                           IF (#temp16ParameterCMAddress <> 255) AND (#temp16ParameterCMAddress >= #NUMBER_OF_CONTROLMODULES_MIN) AND (#temp16ParameterCMAddress <= #NUMBER_OF_CONTROLMODULES)
                               AND (#temp16ParameterType >= #TYPE_NONE) AND (#temp16ParameterType <= #TYPE_STRING) THEN
                               #temp16TempInt1 := #temp16ParameterCMAddress / 32;    //DWORD - Adress
                               #temp16TempInt2 := #temp16ParameterCMAddress MOD 32;  //Bit - Adress
                               //If parameter is forced (FRC) --> Parameter is used
                               IF (((#tempUsed[#temp16TempInt1] AND SHL(IN := #temp32TempDword1, N := INT_TO_UINT(#temp16TempInt2))) <> 0) = TRUE) THEN
                                   CASE #temp16ParameterType OF
                                           // Check of mode is done in satellite blocks
                                       #TYPE_ANALOG:
                                           REGION Analog
                                               //Bit Masking funtionality for calculate the used Analog parameter and Position of the Parameter name in the HMI Text List 
                                               #ProcessInValueType.IndexAnalog := #ProcessInValueType.IndexAnalog OR SHL(IN := #temp32TempDword1, N := INT_TO_UINT(#temp16IndexOfDefinitionProcessIn));
                                               #ProcessInValueType.NameIndexAnalog := #ProcessInValueType.NameIndexAnalog OR SHL(IN := #temp32TempDword1, N := INT_TO_UINT(#temp16IndexOfDefinition));
                                               IF ((#temp16IndexIO >= #PROCESS_VALUES_IN_MIN) AND (#temp16IndexIO <= #PROCESS_VALUES_IN_ANALOG_MAX)) THEN
                                                   //WinCC Parameter View Faceplate logic
                                                   #ProcessInAna[#temp16IndexAnalog].WQC := #ProcessValueInAnalog[#temp16IndexMTP].WQC;
                                                   #ProcessInAna[#temp16IndexAnalog].OSLevel := #ProcessValueInAnalog[#temp16IndexMTP].OSLevel;
                                                   #ProcessInAna[#temp16IndexAnalog].V := #ProcessValueInAnalog[#temp16IndexMTP].V;
                                                   #ProcessInAna[#temp16IndexAnalog].VQC := #ProcessValueInAnalog[#temp16IndexMTP].VQC;
                                                   #ProcessInAna[#temp16IndexAnalog].SclMinCur := #ProcessValueInAnalog[#temp16IndexMTP].SclMinCur;
                                                   #ProcessInAna[#temp16IndexAnalog].SclMaxCur := #ProcessValueInAnalog[#temp16IndexMTP].SclMaxCur;
                                                   #ProcessInAna[#temp16IndexAnalog].UnitCur := #ProcessValueInAnalog[#temp16IndexMTP].UnitCur;
                                                   #ProcessInAna[#temp16IndexAnalog].SclMinExt := #ProcessValueInAnalog[#temp16IndexMTP].SclMinExt;
                                                   #ProcessInAna[#temp16IndexAnalog].SclMaxExt := #ProcessValueInAnalog[#temp16IndexMTP].SclMaxExt;
                                                   #ProcessInAna[#temp16IndexAnalog].UnitExt := #ProcessValueInAnalog[#temp16IndexMTP].UnitExt;
                                                   #ProcessInAna[#temp16IndexAnalog].Apply := #ProcessValueInAnalog[#temp16IndexMTP].Apply;
                                                   #ProcessInAna[#temp16IndexAnalog].ApplyEn := #ProcessValueInAnalog[#temp16IndexMTP].ApplyEn;
                                               END_IF;
                                               #temp16IndexAnalog := #temp16IndexAnalog + 1;
                                           END_REGION
                                       #TYPE_DIGITAL:
                                           REGION Digital
                                               //Bit Masking funtionality for calculate the used Digital parameter and Position of the Parameter name in the HMI Text List 
                                               #ProcessInValueType.IndexDigital := #ProcessInValueType.IndexDigital OR SHL(IN := #temp32TempDword1, N := INT_TO_UINT(#temp16IndexOfDefinitionProcessIn));
                                               #ProcessInValueType.NameIndexDigital := #ProcessInValueType.NameIndexDigital OR SHL(IN := #temp32TempDword1, N := INT_TO_UINT(#temp16IndexOfDefinition));
                                               IF ((#temp16IndexIO >= #PROCESS_VALUES_IN_MIN) AND (#temp16IndexIO <= #PROCESS_VALUES_IN_DIGITAL_MAX)) THEN
                                                   //WinCC Parameter View Faceplate logic
                                                   #ProcessInDint[#temp16IndexDigital].WQC := #ProcessValueInDigital[#temp16IndexMTP].WQC;
                                                   #ProcessInDint[#temp16IndexDigital].OSLevel := #ProcessValueInDigital[#temp16IndexMTP].OSLevel;
                                                   #ProcessInDint[#temp16IndexDigital].V := #ProcessValueInDigital[#temp16IndexMTP].V;
                                                   #ProcessInDint[#temp16IndexDigital].VQC := #ProcessValueInDigital[#temp16IndexMTP].VQC;
                                                   #ProcessInDint[#temp16IndexDigital].SclMinCur := #ProcessValueInDigital[#temp16IndexMTP].SclMinCur;
                                                   #ProcessInDint[#temp16IndexDigital].SclMaxCur := #ProcessValueInDigital[#temp16IndexMTP].SclMaxCur;
                                                   #ProcessInDint[#temp16IndexDigital].UnitCur := #ProcessValueInDigital[#temp16IndexMTP].UnitCur;
                                                   #ProcessInDint[#temp16IndexDigital].SclMinExt := #ProcessValueInDigital[#temp16IndexMTP].SclMinExt;
                                                   #ProcessInDint[#temp16IndexDigital].SclMaxExt := #ProcessValueInDigital[#temp16IndexMTP].SclMaxExt;
                                                   #ProcessInDint[#temp16IndexDigital].UnitExt := #ProcessValueInDigital[#temp16IndexMTP].UnitExt;
                                                   #ProcessInDint[#temp16IndexDigital].Apply := #ProcessValueInDigital[#temp16IndexMTP].Apply;
                                                   #ProcessInDint[#temp16IndexDigital].ApplyEn := #ProcessValueInDigital[#temp16IndexMTP].ApplyEn;
                                               END_IF;
                                               #temp16IndexDigital := #temp16IndexDigital + 1;
                                           END_REGION
                                       #TYPE_BINARY:
                                           REGION Binary
                                               //Bit Masking funtionality for calculate the used Binary parameter and Position of the Parameter name in the HMI Text List 
                                               #ProcessInValueType.IndexBinary := #ProcessInValueType.IndexBinary OR SHL(IN := #temp32TempDword1, N := INT_TO_UINT(#temp16IndexOfDefinitionProcessIn));
                                               #ProcessInValueType.NameIndexBinary := #ProcessInValueType.NameIndexBinary OR SHL(IN := #temp32TempDword1, N := INT_TO_UINT(#temp16IndexOfDefinition));
                                               IF ((#temp16IndexIO >= #PROCESS_VALUES_IN_MIN) AND (#temp16IndexIO <= #PROCESS_VALUES_IN_BINARY_MAX)) THEN
                                                   //WinCC Parameter View Faceplate logic
                                                   #ProcessInBin[#temp16IndexBinary].WQC := #ProcessValueInBinary[#temp16IndexMTP].WQC;
                                                   #ProcessInBin[#temp16IndexBinary].V := #ProcessValueInBinary[#temp16IndexMTP].V;
                                                   #ProcessInBin[#temp16IndexBinary].VQC := #ProcessValueInBinary[#temp16IndexMTP].VQC;
                                                   #ProcessInBin[#temp16IndexBinary].VState0 := #ProcessValueInBinary[#temp16IndexMTP].VState0;
                                                   #ProcessInBin[#temp16IndexBinary].VState1 := #ProcessValueInBinary[#temp16IndexMTP].VState1;
                                               END_IF;
                                               #temp16IndexBinary := #temp16IndexBinary + 1;
                                           END_REGION
                                       #TYPE_STRING:
                                           REGION String
                                               //Bit Masking funtionality for calculate the used String parameter and Position of the Parameter name in the HMI Text List 
                                               #ProcessInValueType.IndexString := #ProcessInValueType.IndexString OR SHL(IN := #temp32TempDword1, N := INT_TO_UINT(#temp16IndexOfDefinitionProcessIn));
                                               #ProcessInValueType.NameIndexString := #ProcessInValueType.NameIndexString OR SHL(IN := #temp32TempDword1, N := INT_TO_UINT(#temp16IndexOfDefinition));
                                               IF ((#temp16IndexIO >= #PROCESS_VALUES_IN_MIN) AND (#temp16IndexIO <= #PROCESS_VALUES_IN_STRING_MAX)) THEN
                                                   //WinCC Parameter View Faceplate logic
                                                   #ProcessInString[#temp16IndexString].WQC := #ProcessValueInString[#temp16IndexMTP].WQC;
                                                   #ProcessInString[#temp16IndexString].V := #ProcessValueInString[#temp16IndexMTP].V;
                                                   #ProcessInString[#temp16IndexString].VQC := #ProcessValueInString[#temp16IndexMTP].VQC;
                                               END_IF;
                                               #temp16IndexString := #temp16IndexString + 1;
                                           END_REGION
                                   END_CASE;
                               END_IF;
                           END_IF;
                           #temp16IndexOfDefinitionProcessIn := #temp16IndexOfDefinitionProcessIn + 1;
                       END_IF;
                   END_FOR;
               END_IF;
           END_IF;
       END_REGION

       REGION Process Out Values

           REGION Get Start and End index details of the Current /Prepared procedure
               //Current/Prepared procedure selection for parameter display in the faceplate
               //#stat32PrecedureProcessOutMap := -1;
               IF NOT (#ProcessOutValueType.ProcedureReqCurInd) THEN
                   #stat32PrecedureProcessOutMap := #tempSetup.procedure.procedure[#stat16ProceCurIndex].ProcedureProcessOutMap[0];
               ELSIF (#ProcessOutValueType.ProcedureReqCurInd) THEN
                   #stat32PrecedureProcessOutMap := #tempSetup.procedure.procedure[#stat16ProceReqIndex].ProcedureProcessOutMap[0];
               END_IF;
           END_REGION
           //Initialize the used variable values          
           #temp32TempDword1 := 16#1;
           #temp16IndexAnalog := 16#0;
           #temp16IndexDigital := 16#0;
           #temp16IndexBinary := 16#0;
           #temp16IndexString := 16#0;
           //Initialize the Process Out Value index and Name index while changing of Procedure and changing of screen selection b/w Prepared and Current procedure
           IF ((#statLasProcedureCur <> #ProcedureCur) OR (#statLasProcedureReq <> #ProcedureReq) OR (#StatLastProceselProcessOut <> #ProcessOutValueType.ProcedureReqCurInd)
               OR (((#ProcedureCur = 16#0) AND NOT #ProcessOutValueType.ProcedureReqCurInd) OR ((#ProcedureReq = 16#0) AND #ProcessOutValueType.ProcedureReqCurInd))) THEN
               #ProcessOutValueType.IndexAnalog := 16#0;
               #ProcessOutValueType.NameIndexAnalog := 16#0;
               #ProcessOutValueType.IndexDigital := 16#0;
               #ProcessOutValueType.NameIndexDigital := 16#0;
               #ProcessOutValueType.IndexBinary := 16#0;
               #ProcessOutValueType.NameIndexBinary := 16#0;
               #ProcessOutValueType.IndexString := 16#0;
               #ProcessOutValueType.NameIndexString := 16#0;
           END_IF;
           //Used/Mapped parameter count with individual parameter type will written from the Tool
           #statTotalProcessOutValues := #MAPPED_PROCESS_OUT_ANALOG + #MAPPED_PROCESS_OUT_DIGITAL + #MAPPED_PROCESS_OUT_BINARY + #MAPPED_PROCESS_OUT_STRING - 1;
           IF (((#ProcedureCur <> 16#0) AND NOT #ProcessOutValueType.ProcedureReqCurInd) OR ((#ProcedureReq <> 16#0) AND #ProcessOutValueType.ProcedureReqCurInd)) THEN
               IF ((#statTotalProcessOutValues >= 0) AND (#statTotalProcessOutValues <= #PROCESS_VALUES_OUT_MAX)) THEN
                   #temp16IndexOfDefinitionProcessOut := 16#0;
                   FOR #temp16IndexOfDefinition := #PROCESS_VALUES_OUT_MIN TO #statTotalProcessOutValues BY 1 DO
                       #temp16ParameterCMAddress := BYTE_TO_INT(#tempSetup.processValueOutData.definition[#temp16IndexOfDefinition].controlModule);
                       #temp16ParameterType := #tempSetup.processValueOutData.definition[#temp16IndexOfDefinition].type;
                       #temp16IndexMTP := #tempSetup.processValueOutData.definition[#temp16IndexOfDefinition].indexMTP;
                       #tempUsed := #tempSetup.processValueOutData.used;
                       // Find the procedure information assigned with the processOut values
                       IF (((#stat32PrecedureProcessOutMap AND SHL(IN := #temp32TempDword1, N := INT_TO_UINT(#temp16IndexOfDefinition))) <> 0) = TRUE) THEN
                           #temp16IndexIO := #tempSetup.processValueOutData.definition[#temp16IndexOfDefinition].indexIO;

                           IF (#temp16ParameterCMAddress <> 255) AND (#temp16ParameterCMAddress >= #NUMBER_OF_CONTROLMODULES_MIN) AND (#temp16ParameterCMAddress <= #NUMBER_OF_CONTROLMODULES)
                               AND (#temp16ParameterType >= #TYPE_NONE) AND (#temp16ParameterType <= #TYPE_STRING) THEN
                               #temp16TempInt1 := #temp16ParameterCMAddress / 32;    //DWORD - Adress
                               #temp16TempInt2 := #temp16ParameterCMAddress MOD 32;  //Bit - Adress
                               //If parameter is forced (FRC) --> Parameter is used
                               IF (((#tempUsed[#temp16TempInt1] AND SHL(IN := #temp32TempDword1, N := INT_TO_UINT(#temp16TempInt2))) <> 0) = TRUE) THEN
                                   CASE #temp16ParameterType OF
                                       #TYPE_ANALOG:
                                           REGION Analog
                                               //Bit Masking funtionality for calculate the used Analog parameter and Position of the Parameter name in the HMI Text List                                         
                                               #ProcessOutValueType.IndexAnalog := #ProcessOutValueType.IndexAnalog OR SHL(IN := #temp32TempDword1, N := INT_TO_UINT(#temp16IndexOfDefinitionProcessOut));
                                               #ProcessOutValueType.NameIndexAnalog := #ProcessOutValueType.NameIndexAnalog OR SHL(IN := #temp32TempDword1, N := INT_TO_UINT(#temp16IndexOfDefinition));
                                               IF ((#temp16IndexIO >= #PROCESS_VALUES_OUT_MIN) AND (#temp16IndexIO <= #PROCESS_VALUES_OUT_ANALOG_MAX)) THEN
                                                   //WinCC Parameter View Faceplate logic
                                                   #ProcessOutAna[#temp16IndexAnalog].WQC := #ProcessValueOutAnalog[#temp16IndexMTP].WQC;
                                                   #ProcessOutAna[#temp16IndexAnalog].V := #ProcessValueOutAnalog[#temp16IndexMTP].V;
                                                   #ProcessOutAna[#temp16IndexAnalog].VSclMin := #ProcessValueOutAnalog[#temp16IndexMTP].VSclMin;
                                                   #ProcessOutAna[#temp16IndexAnalog].VSclMax := #ProcessValueOutAnalog[#temp16IndexMTP].VSclMax;
                                                   #ProcessOutAna[#temp16IndexAnalog].VUnit := #ProcessValueOutAnalog[#temp16IndexMTP].VUnit;
                                               END_IF;
                                               #temp16IndexAnalog := #temp16IndexAnalog + 1;
                                           END_REGION
                                       #TYPE_DIGITAL:
                                           REGION Digital
                                               //Bit Masking funtionality for calculate the used Digital parameter and Position of the Parameter name in the HMI Text List                                         
                                               #ProcessOutValueType.IndexDigital := #ProcessOutValueType.IndexDigital OR SHL(IN := #temp32TempDword1, N := INT_TO_UINT(#temp16IndexOfDefinitionProcessOut));
                                               #ProcessOutValueType.NameIndexDigital := #ProcessOutValueType.NameIndexDigital OR SHL(IN := #temp32TempDword1, N := INT_TO_UINT(#temp16IndexOfDefinition));
                                               IF ((#temp16IndexIO >= #PROCESS_VALUES_OUT_MIN) AND (#temp16IndexIO <= #PROCESS_VALUES_OUT_DIGITAL_MAX)) THEN
                                                   //WinCC Parameter View Faceplate logic
                                                   #ProcessOutDint[#temp16IndexDigital].WQC := #ProcessValueOutDigital[#temp16IndexMTP].WQC;
                                                   #ProcessOutDint[#temp16IndexDigital].V := #ProcessValueOutDigital[#temp16IndexMTP].V;
                                                   #ProcessOutDint[#temp16IndexDigital].VSclMin := #ProcessValueOutDigital[#temp16IndexMTP].VSclMin;
                                                   #ProcessOutDint[#temp16IndexDigital].VSclMax := #ProcessValueOutDigital[#temp16IndexMTP].VSclMax;
                                                   #ProcessOutDint[#temp16IndexDigital].VUnit := #ProcessValueOutDigital[#temp16IndexMTP].VUnit;
                                               END_IF;
                                               #temp16IndexDigital := #temp16IndexDigital + 1;
                                           END_REGION
                                       #TYPE_BINARY:
                                           REGION Binary
                                               //Bit Masking funtionality for calculate the used Binary parameter and Position of the Parameter name in the HMI Text List 
                                               #ProcessOutValueType.IndexBinary := #ProcessOutValueType.IndexBinary OR SHL(IN := #temp32TempDword1, N := INT_TO_UINT(#temp16IndexOfDefinitionProcessOut));
                                               #ProcessOutValueType.NameIndexBinary := #ProcessOutValueType.NameIndexBinary OR SHL(IN := #temp32TempDword1, N := INT_TO_UINT(#temp16IndexOfDefinition));
                                               IF ((#temp16IndexIO >= #PROCESS_VALUES_OUT_MIN) AND (#temp16IndexIO <= #PROCESS_VALUES_OUT_BINARY_MAX)) THEN
                                                   //WinCC Parameter View Faceplate logic
                                                   #ProcessOutBin[#temp16IndexBinary].WQC := #ProcessValueOutBinary[#temp16IndexMTP].WQC;
                                                   #ProcessOutBin[#temp16IndexBinary].V := #ProcessValueOutBinary[#temp16IndexMTP].V;
                                                   #ProcessOutBin[#temp16IndexBinary].VState0 := #ProcessValueOutBinary[#temp16IndexMTP].VState0;
                                                   #ProcessOutBin[#temp16IndexBinary].VState1 := #ProcessValueOutBinary[#temp16IndexMTP].VState1;
                                               END_IF;
                                               #temp16IndexBinary := #temp16IndexBinary + 1;
                                           END_REGION
                                       #TYPE_STRING:
                                           REGION String
                                               //Bit Masking funtionality for calculate the used String parameter and Position of the Parameter name in the HMI Text List 
                                               #ProcessOutValueType.IndexString := #ProcessOutValueType.IndexString OR SHL(IN := #temp32TempDword1, N := INT_TO_UINT(#temp16IndexOfDefinitionProcessOut));
                                               #ProcessOutValueType.NameIndexString := #ProcessOutValueType.NameIndexString OR SHL(IN := #temp32TempDword1, N := INT_TO_UINT(#temp16IndexOfDefinition));
                                               IF ((#temp16IndexIO >= #PROCESS_VALUES_OUT_MIN) AND (#temp16IndexIO <= #PROCESS_VALUES_OUT_STRING_MAX)) THEN
                                                   //WinCC Parameter View Faceplate logic
                                                   #ProcessOutString[#temp16IndexString].WQC := #ProcessValueOutString[#temp16IndexMTP].WQC;
                                                   #ProcessOutString[#temp16IndexString].Text := #ProcessValueOutString[#temp16IndexMTP].Text;
                                               END_IF;
                                               #temp16IndexString := #temp16IndexString + 1;
                                           END_REGION
                                   END_CASE;
                               END_IF;
                           END_IF;
                           #temp16IndexOfDefinitionProcessOut := #temp16IndexOfDefinitionProcessOut + 1;
                       END_IF;
                   END_FOR;
               END_IF;
           END_IF;
       END_REGION

       REGION Report Values

           REGION Get Start and End index details of the Current /Prepared procedure
               //Current/Prepared procedure selection for parameter display in the faceplate
              // #stat32PrecedureReportMap := -1;
               IF NOT (#ReportValueType.ProcedureReqCurInd) THEN
                   #stat32PrecedureReportMap := #tempSetup.procedure.procedure[#stat16ProceCurIndex].ProcedureReportMap[0];
               ELSIF (#ReportValueType.ProcedureReqCurInd) THEN
                   #stat32PrecedureReportMap := #tempSetup.procedure.procedure[#stat16ProceReqIndex].ProcedureReportMap[0];
               END_IF;
           END_REGION
           //Initialize the used variable values        
           #temp32TempDword1 := 16#1;
           #temp16IndexAnalog := 16#0;
           #temp16IndexDigital := 16#0;
           #temp16IndexBinary := 16#0;
           #temp16IndexString := 16#0;
           //Initialize the Process Out Value index and Name index while changing of Procedure and changing of screen selection b/w Prepared and Current procedure
           IF ((#statLasProcedureCur <> #ProcedureCur) OR (#statLasProcedureReq <> #ProcedureReq) OR (#StatLastProceselReport <> #ReportValueType.ProcedureReqCurInd)
               OR (((#ProcedureCur = 16#0) AND NOT #ReportValueType.ProcedureReqCurInd) OR ((#ProcedureReq = 16#0) AND #ReportValueType.ProcedureReqCurInd))) THEN
               #ReportValueType.IndexAnalog := 16#0;
               #ReportValueType.NameIndexAnalog := 16#0;
               #ReportValueType.IndexDigital := 16#0;
               #ReportValueType.NameIndexDigital := 16#0;
               #ReportValueType.IndexBinary := 16#0;
               #ReportValueType.NameIndexBinary := 16#0;
               #ReportValueType.IndexString := 16#0;
               #ReportValueType.NameIndexString := 16#0;
           END_IF;
           //Used/Mapped parameter count with individual parameter type will written from the Tool
           #statTotalReportValues := #MAPPED_REPORT_ANALOG + #MAPPED_REPORT_DIGITAL + #MAPPED_REPORT_BINARY + #MAPPED_REPORT_STRING - 1;
           IF (((#ProcedureCur <> 16#0) AND NOT #ReportValueType.ProcedureReqCurInd) OR ((#ProcedureReq <> 16#0) AND #ReportValueType.ProcedureReqCurInd)) THEN
               IF ((#statTotalReportValues >= 0) AND (#statTotalReportValues <= #REPORT_VALUES_MAX)) THEN
                   #temp16IndexOfDefinitionReport := 16#0;
                   FOR #temp16IndexOfDefinition := #REPORT_VALUES_MIN TO #statTotalReportValues BY 1 DO
                       #temp16ParameterCMAddress := BYTE_TO_INT(#tempSetup.reportValueData.definition[#temp16IndexOfDefinition].controlModule);
                       #temp16ParameterType := #tempSetup.reportValueData.definition[#temp16IndexOfDefinition].type;
                       #temp16IndexMTP := #tempSetup.reportValueData.definition[#temp16IndexOfDefinition].indexMTP;
                       #tempUsed := #tempSetup.reportValueData.used;
                       // Find the procedure information assigned with the report values
                       IF (((#stat32PrecedureReportMap AND SHL(IN := #temp32TempDword1, N := INT_TO_UINT(#temp16IndexOfDefinition))) <> 0) = TRUE) THEN
                           #temp16IndexIO := #tempSetup.reportValueData.definition[#temp16IndexOfDefinition].indexIO;

                           IF (#temp16ParameterCMAddress <> 255) AND (#temp16ParameterCMAddress >= #NUMBER_OF_CONTROLMODULES_MIN) AND (#temp16ParameterCMAddress <= #NUMBER_OF_CONTROLMODULES)
                               AND (#temp16ParameterType >= #TYPE_NONE) AND (#temp16ParameterType <= #TYPE_STRING) THEN
                               #temp16TempInt1 := #temp16ParameterCMAddress / 32;    //DWORD - Adress
                               #temp16TempInt2 := #temp16ParameterCMAddress MOD 32;  //Bit - Adress
                               //If parameter is forced (FRC) --> Parameter is used
                               IF (((#tempUsed[#temp16TempInt1] AND SHL(IN := #temp32TempDword1, N := INT_TO_UINT(#temp16TempInt2))) <> 0) = TRUE) THEN
                                   CASE #temp16ParameterType OF
                                       #TYPE_ANALOG:
                                           REGION Analog
                                               //Bit Masking funtionality for calculate the used Analog parameter and Position of the Parameter name in the HMI Text List 
                                               #ReportValueType.IndexAnalog := #ReportValueType.IndexAnalog OR SHL(IN := #temp32TempDword1, N := INT_TO_UINT(#temp16IndexOfDefinitionReport));
                                               #ReportValueType.NameIndexAnalog := #ReportValueType.NameIndexAnalog OR SHL(IN := #temp32TempDword1, N := INT_TO_UINT(#temp16IndexOfDefinition));
                                               IF ((#temp16IndexIO >= #REPORT_VALUES_MIN) AND (#temp16IndexIO <= #REPORT_VALUES_ANALOG_MAX)) THEN
                                                   //WinCC Parameter View Faceplate logic
                                                   #ReportAna[#temp16IndexAnalog].WQC := #ReportValueAnalog[#temp16IndexMTP].WQC;
                                                   #ReportAna[#temp16IndexAnalog].V := #ReportValueAnalog[#temp16IndexMTP].V;
                                                   #ReportAna[#temp16IndexAnalog].VSclMin := #ReportValueAnalog[#temp16IndexMTP].VSclMin;
                                                   #ReportAna[#temp16IndexAnalog].VSclMax := #ReportValueAnalog[#temp16IndexMTP].VSclMax;
                                                   #ReportAna[#temp16IndexAnalog].VUnit := #ReportValueAnalog[#temp16IndexMTP].VUnit;
                                                   #ReportAna[#temp16IndexAnalog].MissedValue := #ReportValueAnalog[#temp16IndexMTP].MissedValue;
                                               END_IF;
                                               #temp16IndexAnalog := #temp16IndexAnalog + 1;
                                           END_REGION
                                       #TYPE_DIGITAL:
                                           REGION Digital
                                               //Bit Masking funtionality for calculate the used Digital parameter and Position of the Parameter name in the HMI Text List 
                                               #ReportValueType.IndexDigital := #ReportValueType.IndexDigital OR SHL(IN := #temp32TempDword1, N := INT_TO_UINT(#temp16IndexOfDefinitionReport));
                                               #ReportValueType.NameIndexDigital := #ReportValueType.NameIndexDigital OR SHL(IN := #temp32TempDword1, N := INT_TO_UINT(#temp16IndexOfDefinition));
                                               IF ((#temp16IndexIO >= #REPORT_VALUES_MIN) AND (#temp16IndexIO <= #REPORT_VALUES_DIGITAL_MAX)) THEN
                                                   //WinCC Parameter View Faceplate logic
                                                   #ReportDint[#temp16IndexDigital].WQC := #ReportValueDigital[#temp16IndexMTP].WQC;
                                                   #ReportDint[#temp16IndexDigital].V := #ReportValueDigital[#temp16IndexMTP].V;
                                                   #ReportDint[#temp16IndexDigital].VSclMin := #ReportValueDigital[#temp16IndexMTP].VSclMin;
                                                   #ReportDint[#temp16IndexDigital].VSclMax := #ReportValueDigital[#temp16IndexMTP].VSclMax;
                                                   #ReportDint[#temp16IndexDigital].VUnit := #ReportValueDigital[#temp16IndexMTP].VUnit;
                                                   #ReportDint[#temp16IndexDigital].MissedValue := #ReportValueDigital[#temp16IndexMTP].MissedValue;
                                               END_IF;
                                               #temp16IndexDigital := #temp16IndexDigital + 1;
                                           END_REGION
                                       #TYPE_BINARY:
                                           REGION Binary
                                               //Bit Masking funtionality for calculate the used Binary parameter and Position of the Parameter name in the HMI Text List 
                                               #ReportValueType.IndexBinary := #ReportValueType.IndexBinary OR SHL(IN := #temp32TempDword1, N := INT_TO_UINT(#temp16IndexOfDefinitionReport));
                                               #ReportValueType.NameIndexBinary := #ReportValueType.NameIndexBinary OR SHL(IN := #temp32TempDword1, N := INT_TO_UINT(#temp16IndexOfDefinition));
                                               IF ((#temp16IndexIO >= #REPORT_VALUES_MIN) AND (#temp16IndexIO <= #REPORT_VALUES_BINARY_MAX)) THEN
                                                   //WinCC Parameter View Faceplate logic
                                                   #ReportBin[#temp16IndexBinary].WQC := #ReportValueBinary[#temp16IndexMTP].WQC;
                                                   #ReportBin[#temp16IndexBinary].V := #ReportValueBinary[#temp16IndexMTP].V;
                                                   #ReportBin[#temp16IndexBinary].VState0 := #ReportValueBinary[#temp16IndexMTP].VState0;
                                                   #ReportBin[#temp16IndexBinary].VState1 := #ReportValueBinary[#temp16IndexMTP].VState1;
                                                   #ReportBin[#temp16IndexBinary].MissedValue := #ReportValueBinary[#temp16IndexMTP].MissedValue;
                                               END_IF;
                                               #temp16IndexBinary := #temp16IndexBinary + 1;
                                           END_REGION
                                       #TYPE_STRING:
                                           REGION String
                                               //Bit Masking funtionality for calculate the used String parameter and Position of the Parameter name in the HMI Text List 
                                               #ReportValueType.IndexString := #ReportValueType.IndexString OR SHL(IN := #temp32TempDword1, N := INT_TO_UINT(#temp16IndexOfDefinitionReport));
                                               #ReportValueType.NameIndexString := #ReportValueType.NameIndexString OR SHL(IN := #temp32TempDword1, N := INT_TO_UINT(#temp16IndexOfDefinition));
                                               IF ((#temp16IndexIO >= #REPORT_VALUES_MIN) AND (#temp16IndexIO <= #REPORT_VALUES_STRING_MAX)) THEN

                                                   //WinCC Parameter View Faceplate logic
                                                   #ReportString[#temp16IndexString].WQC := #ReportValueString[#temp16IndexMTP].WQC;
                                                   #ReportString[#temp16IndexString].Text := #ReportValueString[#temp16IndexMTP].Text;
                                                   #ReportString[#temp16IndexString].MissedValue := #ReportValueString[#temp16IndexMTP].MissedValue;
                                               END_IF;
                                               #temp16IndexString := #temp16IndexString + 1;
                                           END_REGION
                                   END_CASE;
                               END_IF;
                           END_IF;
                           #temp16IndexOfDefinitionReport := #temp16IndexOfDefinitionReport + 1;
                       END_IF;
                   END_FOR;
               END_IF;
           END_IF;
       END_REGION  

       //Move last valid value 
       #statLasProcedureCur := #ProcedureCur;
       #statLasProcedureReq := #ProcedureReq;
       #statLastReqProcedSelected := #ProcedureParaType.ProcedureReqCurInd;
       #StatLastProceselProcessIn := #ProcessInValueType.ProcedureReqCurInd;
       #StatLastProceselProcessOut := #ProcessOutValueType.ProcedureReqCurInd;
       #StatLastProceselReport := #ReportValueType.ProcedureReqCurInd;
END_FUNCTION_BLOCK

FUNCTION_BLOCK "CM_Interface"   // FB5, SCL
{ S7_Optimized_Access := 'TRUE' }
// stored: MemoryReserve 100, SetENOAutomatically false
   VAR_INPUT
      CmCommand { ExternalAccessible := 'False'; ExternalVisible := 'False'; ExternalWritable := 'False'} : Array[0..29] of Bool;
      Procedure_Param { ExternalAccessible := 'False'; ExternalVisible := 'False'; ExternalWritable := 'False'} : Array[0..31] of Real;
      Config_Param : Array[0..31] of Bool;
      ProcessValueIn_Bool : Array[0..31] of Bool;
      ProcessValueIn_Real : Array[0..31] of Real;
      CmFbOnOff { ExternalAccessible := 'False'; ExternalVisible := 'False'; ExternalWritable := 'False'} : Array[0..29] of Bool;
      DosingSpeed : Real;
      Auto_Man : Bool;
      Oos : Bool;
   END_VAR
   VAR_OUTPUT
      CM_P100 { ExternalAccessible := 'False'; ExternalVisible := 'False'; ExternalWritable := 'False'} : "DigVal";
      CM_P101 { ExternalAccessible := 'False'; ExternalVisible := 'False'; ExternalWritable := 'False'} : "DigVal";
      CM_FIC100 { ExternalAccessible := 'False'; ExternalVisible := 'False'; ExternalWritable := 'False'} : "DigVal";
      CM_V100 { ExternalAccessible := 'False'; ExternalVisible := 'False'; ExternalWritable := 'False'} : "DigVal";
      FlowRate { ExternalAccessible := 'False'; ExternalVisible := 'False'; ExternalWritable := 'False'} : "AnaVal";
      Liter { ExternalAccessible := 'False'; ExternalVisible := 'False'; ExternalWritable := 'False'} : "AnaVal";
      ExternalLevel : "AnaVal";
      PEA_inlet_Vlv_opened : "DigVal";
      PVConnected : "DigVal";
   END_VAR
   VAR
      Pos_edge : Bool;
      Neg_edge : Bool;
   END_VAR
   VAR_TEMP
      State : "Service_States";
   END_VAR
BEGIN
   REGION Bool TO DigVal
       //CM Pump 100
       "BoolToDigVal"(In := #CmCommand[0],
                      ST := 16#80,
                      Out => #CM_P100);
       //CM Pump 101
       "BoolToDigVal"(In := #CmCommand[1],
                      ST := 16#80,
                      Out => #CM_P101);
       //CM Controler 100
       "BoolToDigVal"(In := #CmCommand[2],
                      ST := 16#80,
                      Out => #CM_FIC100);
       //CM Valve 100
       "BoolToDigVal"(In := #CmCommand[3],
                      ST := 16#80,
                      Out => #CM_V100);
   END_REGION

   REGION Real TO AnaVal
       //Flow
       "RealToAnaVal"(In := #Procedure_Param[0],
                      ST := 16#80,
                      Out => #FlowRate);
       //Liter
       "RealToAnaVal"(In := #Procedure_Param[1],
                      ST := 16#80,
                      Out => #Liter);
                   END_REGION

   REGION other values
       //Dosing Speed
       "Dose".ProcessValueOutAnalogIn[0] := #DosingSpeed;

       //Configuration parameter
       "BoolToDigVal"(In := #Config_Param[0],
                      ST := 16#80,
                      Out => #PVConnected);
       //process value input
       "RealToAnaVal"(In := #ProcessValueIn_Real[0],
                      ST := 16#80,
                      Out => #ExternalLevel);
       "BoolToDigVal"(In := #ProcessValueIn_Bool[0],
                      ST := 16#80,
                      Out => #PEA_inlet_Vlv_opened);
   END_REGION


   REGION Set auto/man mode & Int/Ext
       //check for positive edge at Dose.Oos
       "R_TRIG_DB"(CLK := #Oos,
                   Q => #Neg_edge);

       //Set POs to auto mode
       IF #Auto_Man = TRUE THEN
           "FIC100_Type".Cmd_Man := FALSE;
           "P100_Type".Cmd_Man := FALSE;
           "V100_Type".Cmd_Man := FALSE;
           "P101_Type".Cmd_Man := FALSE;
           "FIC100_Type".Cmd_Auto := TRUE;
           "P100_Type".Cmd_Auto := TRUE;
           "V100_Type".Cmd_Auto := TRUE;
           "P101_Type".Cmd_Auto := TRUE;
       //Set POs to man mode
       ELSIF #Neg_edge = TRUE THEN
           "FIC100_Type".Cmd_Auto := FALSE;
           "P100_Type".Cmd_Auto := FALSE;
           "V100_Type".Cmd_Auto := FALSE;
           "P101_Type".Cmd_Auto := FALSE;
           "FIC100_Type".Cmd_Man := TRUE;
           "P100_Type".Cmd_Man := TRUE;
           "V100_Type".Cmd_Man := TRUE;
           "P101_Type".Cmd_Man := TRUE;
       //Reset Value
       ELSE
           "FIC100_Type".Cmd_Auto := FALSE;
           "P100_Type".Cmd_Auto := FALSE;
           "V100_Type".Cmd_Auto := FALSE;
           "P101_Type".Cmd_Auto := FALSE;
           "FIC100_Type".Cmd_Man := FALSE;
           "P100_Type".Cmd_Man := FALSE;
           "V100_Type".Cmd_Man := FALSE;
           "P101_Type".Cmd_Man := FALSE;
       END_IF;
   END_REGION
END_FUNCTION_BLOCK

FUNCTION_BLOCK "Service_Command_Logic"   // FB3, SCL
{ S7_Optimized_Access := 'TRUE' }
// stored: MemoryReserve 100, SetENOAutomatically false
   VAR_INPUT
      Level : Real;
      ProcedureID_cur : DWord;
   END_VAR
   VAR_TEMP
      i : Int;
      State : "Service_States";
   END_VAR
BEGIN
   //Set service to hold, if the level of the tank falls under 0,45 during the 
   //procedures DoseByVolume and DoseByFlow
   IF #Level < 45 AND "Dose".Information.state = #State.Execute AND "Dose".MTP.ServiceControl.ProcedureCur <> 3 THEN
       "Dose".CommandForce.hold := TRUE;
       FOR #i := 0 TO 1 BY 1 DO
           "Dose".Procedure[#i].ProcedureEnable.Unhold.ST := 16#80;
           "Dose".Procedure[#i].ProcedureEnable.Unhold.Value := false;
       END_FOR;
   END_IF;
   IF "Dose".Information.state = #State.Held THEN
       "Dose".CommandForce.hold := FALSE;
   END_IF;
   IF "Dose".Information.state = #State.Held AND #Level >= 1.0 THEN
       FOR #i := 0 TO 1 BY 1 DO
           "Dose".Procedure[#i].ProcedureEnable.Unhold.ST := 16#80;
           "Dose".Procedure[#i].ProcedureEnable.Unhold.Value := true;
       END_FOR;
   END_IF;


   //Set service to abort, if the pump is in failure
   IF "P100_Type".GrpErr = True OR "P101_Type".GrpErr THEN
       "Dose".CommandForce.abort := TRUE;
       FOR #i := 0 TO 2 BY 1 DO
           "Dose".Procedure[#i].ProcedureEnable.Start.ST := 16#80;
           "Dose".Procedure[#i].ProcedureEnable.Start.Value := false;
       END_FOR;
   ELSIF ("Dose".Information.state = #State.Aborted OR "Dose".Information.state = #State.Idle) AND ("P100_Type".GrpErr = False OR "P101_Type".GrpErr) THEN
       "Dose".CommandForce.abort := false;
       FOR #i := 0 TO 2 BY 1 DO
           "Dose".Procedure[#i].ProcedureEnable.Start.ST := 16#80;
           "Dose".Procedure[#i].ProcedureEnable.Start.Value := true;
       END_FOR;
   END_IF;
END_FUNCTION_BLOCK

FUNCTION "BoolToDigVal" : Void   // FC10, SCL
{ S7_Optimized_Access := 'TRUE' }
// stored: SetENOAutomatically false
   VAR_INPUT
      In : Bool;
      ST : Byte;
   END_VAR
   VAR_OUTPUT
      Out : "DigVal";
   END_VAR
BEGIN
   #Out.ST := #ST;
   #Out.Value := #In;
END_FUNCTION

FUNCTION "PositionText" : Void   // FC18, SCL
{ S7_Optimized_Access := 'TRUE' }
// stored: SetENOAutomatically false
   VAR_INPUT
      PosID_1 : Bool;
      PosID_2 : Bool;
      PosID_3 : Bool;
      PosID_4 : Bool;
      PosID_5 : Bool;
      PosID_6 : Bool;
      PosID_7 : Bool;
      PosID_8 : Bool;
      PosID_9 : Bool;
      PosID_10 : Bool;
      PosID_0 : Bool;
   END_VAR
BEGIN
   IF #PosID_1 = True THEN
       "Dose".PosTextIDLi := 1;
   ELSIF #PosID_2 = True THEN
       "Dose".PosTextIDLi := 2;
   ELSIF #PosID_3 = True THEN
       "Dose".PosTextIDLi := 3;
   ELSIF #PosID_4 = True THEN
       "Dose".PosTextIDLi := 4;
   ELSIF #PosID_5 = True THEN
       "Dose".PosTextIDLi := 5;
   ELSIF #PosID_6 = True THEN
       "Dose".PosTextIDLi := 6;
   ELSIF #PosID_7 = True THEN
       "Dose".PosTextIDLi := 7;
   ELSIF #PosID_8 = True THEN
       "Dose".PosTextIDLi := 8;
   ELSIF #PosID_9 = True THEN
       "Dose".PosTextIDLi := 9;
   ELSIF #PosID_10 = True THEN
       "Dose".PosTextIDLi := 10;
   ELSIF #PosID_0 = True THEN
       "Dose".PosTextIDLi := 0;
   END_IF;
END_FUNCTION

FUNCTION "FIC100" : Void   // FC5, FBD
{ S7_Optimized_Access := 'TRUE' }
// stored: SetENOAutomatically false
   VAR_TEMP
      Temp : "DigVal";
      State : "Service_States";
      Interlock : "DigVal";
   END_VAR
BEGIN

REGION Network 1: PIDConL interconnections
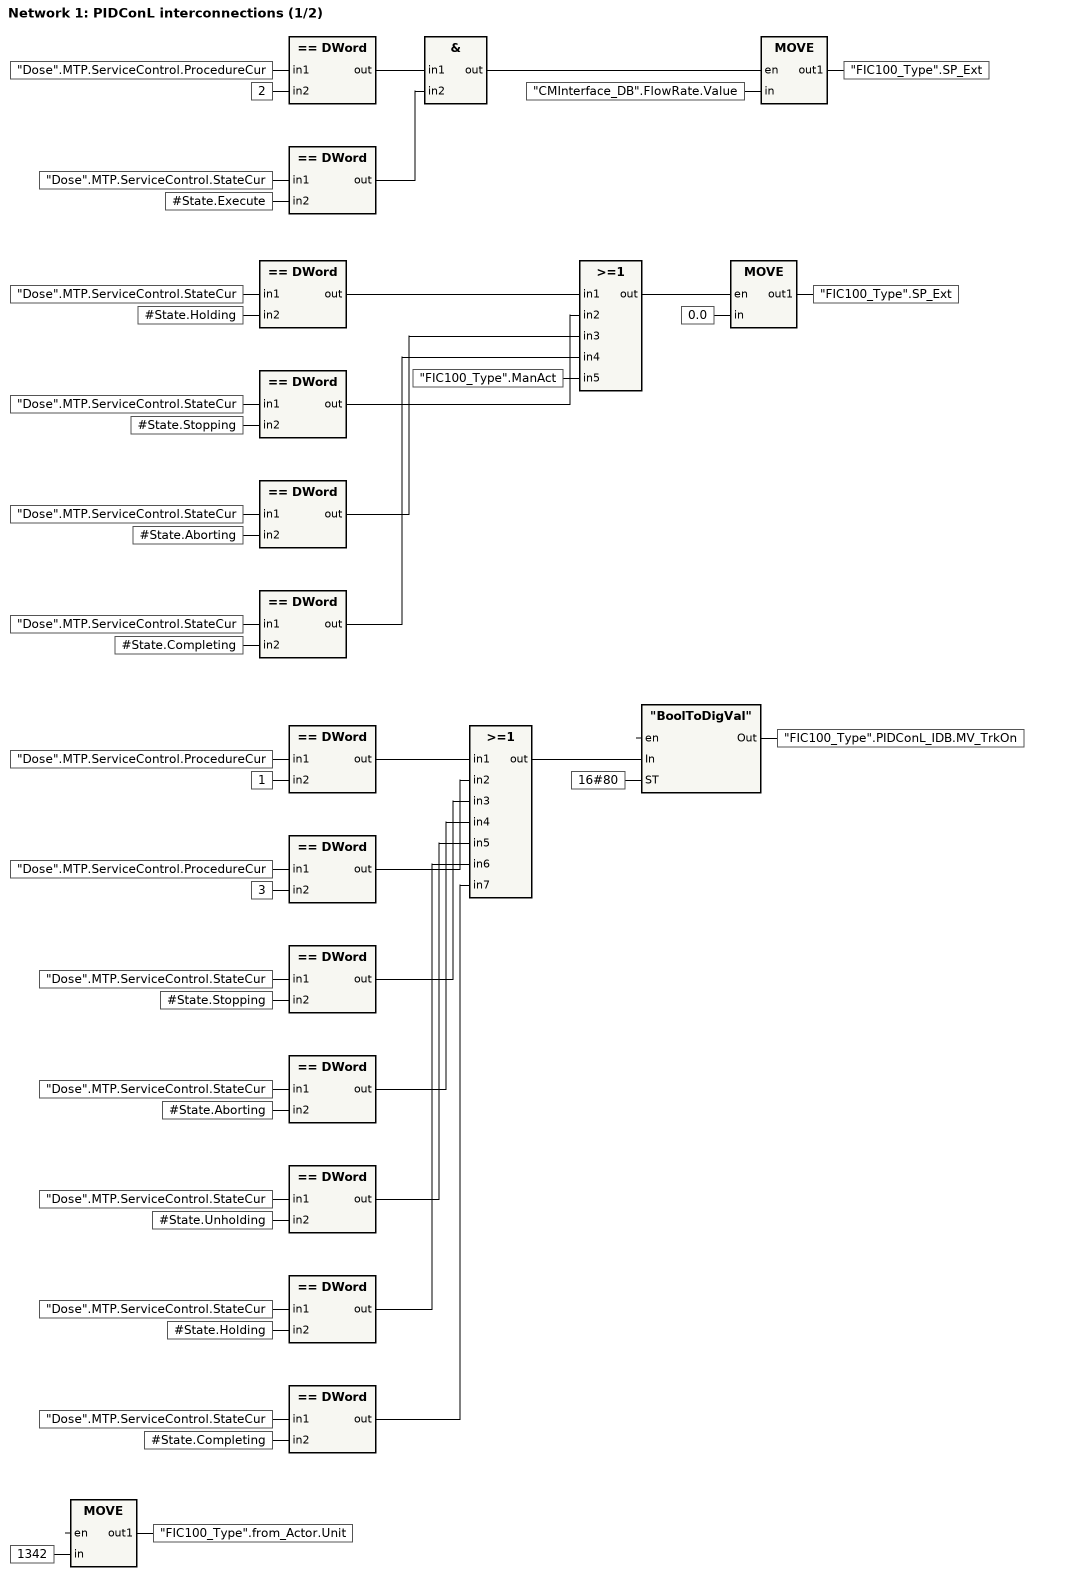
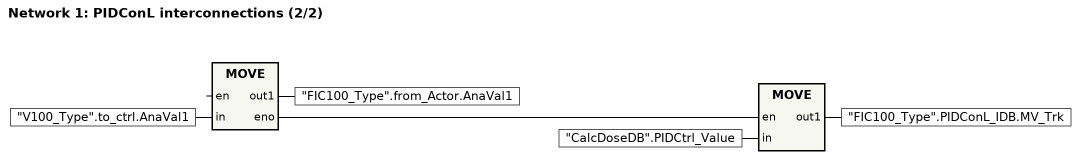
   IF ("Dose".MTP.ServiceControl.ProcedureCur = 2) AND ("Dose".MTP.ServiceControl.StateCur = #State.Execute) THEN
       "FIC100_Type".SP_Ext := "CMInterface_DB".FlowRate.Value;
   END_IF;
   IF ("Dose".MTP.ServiceControl.StateCur = #State.Holding) OR ("Dose".MTP.ServiceControl.StateCur = #State.Stopping) OR ("Dose".MTP.ServiceControl.StateCur = #State.Aborting) OR ("Dose".MTP.ServiceControl.StateCur = #State.Completing) OR "FIC100_Type".ManAct THEN
       "FIC100_Type".SP_Ext := 0.0;
   END_IF;
   "BoolToDigVal"(In := ("Dose".MTP.ServiceControl.ProcedureCur = 1) OR ("Dose".MTP.ServiceControl.ProcedureCur = 3) OR ("Dose".MTP.ServiceControl.StateCur = #State.Stopping) OR ("Dose".MTP.ServiceControl.StateCur = #State.Aborting) OR ("Dose".MTP.ServiceControl.StateCur = #State.Unholding) OR ("Dose".MTP.ServiceControl.StateCur = #State.Holding) OR ("Dose".MTP.ServiceControl.StateCur = #State.Completing),
                  ST := 16#80,
                  Out => "FIC100_Type".PIDConL_IDB.MV_TrkOn);
   "FIC100_Type".from_Actor.Unit := 1342;
   "FIC100_Type".from_Actor.AnaVal1 := "V100_Type".to_ctrl.AnaVal1;
   "FIC100_Type".PIDConL_IDB.MV_Trk := "CalcDoseDB".PIDCtrl_Value;
END_REGION

REGION Network 2: PIDCon
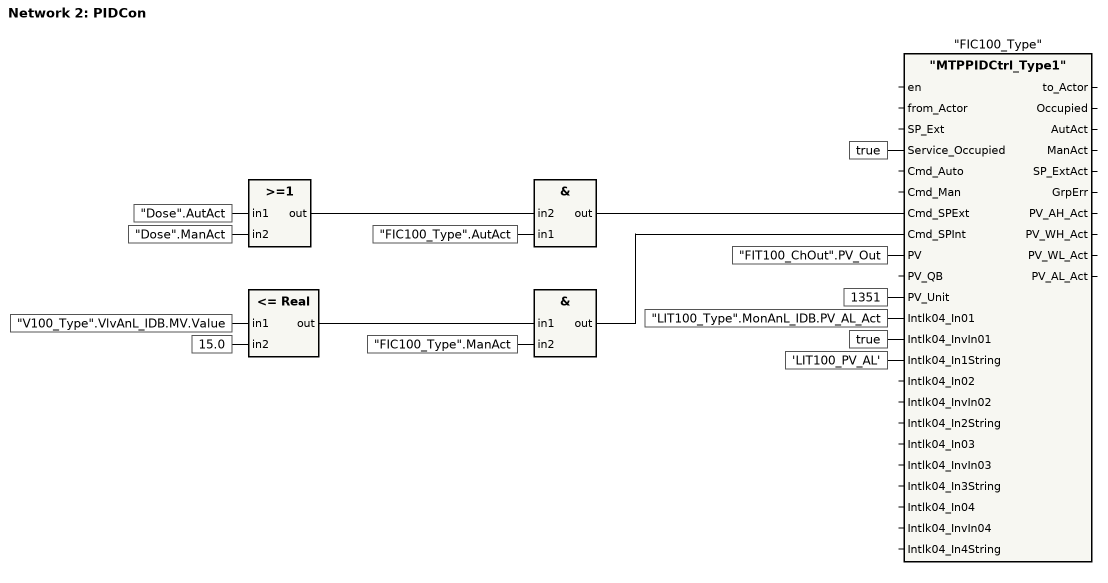
   "FIC100_Type"(Service_Occupied := true,   // "MTPPIDCtrl_Type1"
                 Cmd_SPExt := ("Dose".AutAct OR "Dose".ManAct) AND "FIC100_Type".AutAct,
                 Cmd_SPInt := ("V100_Type".VlvAnL_IDB.MV.Value <= 15.0) AND "FIC100_Type".ManAct,
                 PV := "FIT100_ChOut".PV_Out,
                 PV_Unit := 1351,
                 Intlk04_In01 := "LIT100_Type".MonAnL_IDB.PV_AL_Act,
                 Intlk04_InvIn01 := true,
                 Intlk04_In1String := 'LIT100_PV_AL');
END_REGION
END_FUNCTION

FUNCTION_BLOCK "MTPPIDCtrl_Type1"   // FB14, FBD
{ S7_Optimized_Access := 'TRUE' }
// stored: MemoryReserve 100, SetENOAutomatically false
   VAR_INPUT
      from_Actor { ExternalAccessible := 'False'; ExternalVisible := 'False'; ExternalWritable := 'False'} : "StruCm";
      SP_Ext { ExternalAccessible := 'False'; ExternalVisible := 'False'; ExternalWritable := 'False'} : Real;
      Service_Occupied { ExternalAccessible := 'False'; ExternalVisible := 'False'; ExternalWritable := 'False'} : Bool;
      Cmd_Auto { ExternalAccessible := 'False'; ExternalVisible := 'False'; ExternalWritable := 'False'} : Bool;
      Cmd_Man { ExternalAccessible := 'False'; ExternalVisible := 'False'; ExternalWritable := 'False'} : Bool;
      Cmd_SPExt { ExternalAccessible := 'False'; ExternalVisible := 'False'; ExternalWritable := 'False'} : Bool;
      Cmd_SPInt { ExternalAccessible := 'False'; ExternalVisible := 'False'; ExternalWritable := 'False'} : Bool;
      PV { ExternalAccessible := 'False'; ExternalVisible := 'False'; ExternalWritable := 'False'} : Word;
      PV_QB { ExternalAccessible := 'False'; ExternalVisible := 'False'; ExternalWritable := 'False'} : Bool := true;
      PV_Unit { ExternalAccessible := 'False'; ExternalVisible := 'False'; ExternalWritable := 'False'} : Int := 1342;
      Intlk04_In01 { ExternalAccessible := 'False'; ExternalVisible := 'False'; ExternalWritable := 'False'} : "DigVal";
      Intlk04_InvIn01 { ExternalAccessible := 'False'; ExternalVisible := 'False'; ExternalWritable := 'False'} : Bool;
      Intlk04_In1String : String;
      Intlk04_In02 { ExternalAccessible := 'False'; ExternalVisible := 'False'; ExternalWritable := 'False'} : "DigVal";
      Intlk04_InvIn02 { ExternalAccessible := 'False'; ExternalVisible := 'False'; ExternalWritable := 'False'} : Bool;
      Intlk04_In2String : String;
      Intlk04_In03 { ExternalAccessible := 'False'; ExternalVisible := 'False'; ExternalWritable := 'False'} : "DigVal";
      Intlk04_InvIn03 { ExternalAccessible := 'False'; ExternalVisible := 'False'; ExternalWritable := 'False'} : Bool;
      Intlk04_In3String : String;
      Intlk04_In04 { ExternalAccessible := 'False'; ExternalVisible := 'False'; ExternalWritable := 'False'} : "DigVal";
      Intlk04_InvIn04 { ExternalAccessible := 'False'; ExternalVisible := 'False'; ExternalWritable := 'False'} : Bool;
      Intlk04_In4String : String;
   END_VAR
   VAR_OUTPUT
      to_Actor { ExternalAccessible := 'False'; ExternalVisible := 'False'; ExternalWritable := 'False'} : "StruCm";
      Occupied { ExternalAccessible := 'False'; ExternalVisible := 'False'; ExternalWritable := 'False'} : Bool;   // Occupied by a Service procedure
      AutAct { ExternalAccessible := 'False'; ExternalVisible := 'False'; ExternalWritable := 'False'} : Bool;
      ManAct { ExternalAccessible := 'False'; ExternalVisible := 'False'; ExternalWritable := 'False'} : Bool;
      SP_ExtAct { ExternalAccessible := 'False'; ExternalVisible := 'False'; ExternalWritable := 'False'} : Bool;
      GrpErr { ExternalAccessible := 'False'; ExternalVisible := 'False'; ExternalWritable := 'False'} : Bool;
      PV_AH_Act { ExternalAccessible := 'False'; ExternalVisible := 'False'; ExternalWritable := 'False'} : Bool;
      PV_WH_Act { ExternalAccessible := 'False'; ExternalVisible := 'False'; ExternalWritable := 'False'} : Bool;
      PV_WL_Act { ExternalAccessible := 'False'; ExternalVisible := 'False'; ExternalWritable := 'False'} : Bool;
      PV_AL_Act { ExternalAccessible := 'False'; ExternalVisible := 'False'; ExternalWritable := 'False'} : Bool;
   END_VAR
   VAR
      AnIn_IDB { ExternalAccessible := 'False'; ExternalVisible := 'False'; ExternalWritable := 'False'} : "AnIn";
      Intlk04_IDB : "Intlk04";
      PIDConL_IDB { S7_SetPoint := 'True'} : "PIDConL";
      MTPPIDCtrl_IDB { ExternalVisible := 'False'; S7_SetPoint := 'True'} : "MTPPIDCtrl";
   END_VAR
   VAR_TEMP
      Intlock : "DigVal";
      PV_Out : "AnaVal";
      ScaleOut : "ScaVal";
      BadOut : "DigVal";
      CSF_NOP : "DigVal";
   END_VAR
   // Intlk04_In01.Value := true;
   // Intlk04_In02.Value := true;
   // Intlk04_In03.Value := true;
   // Intlk04_In04.Value := true;
BEGIN

REGION Network 1: Mod switch
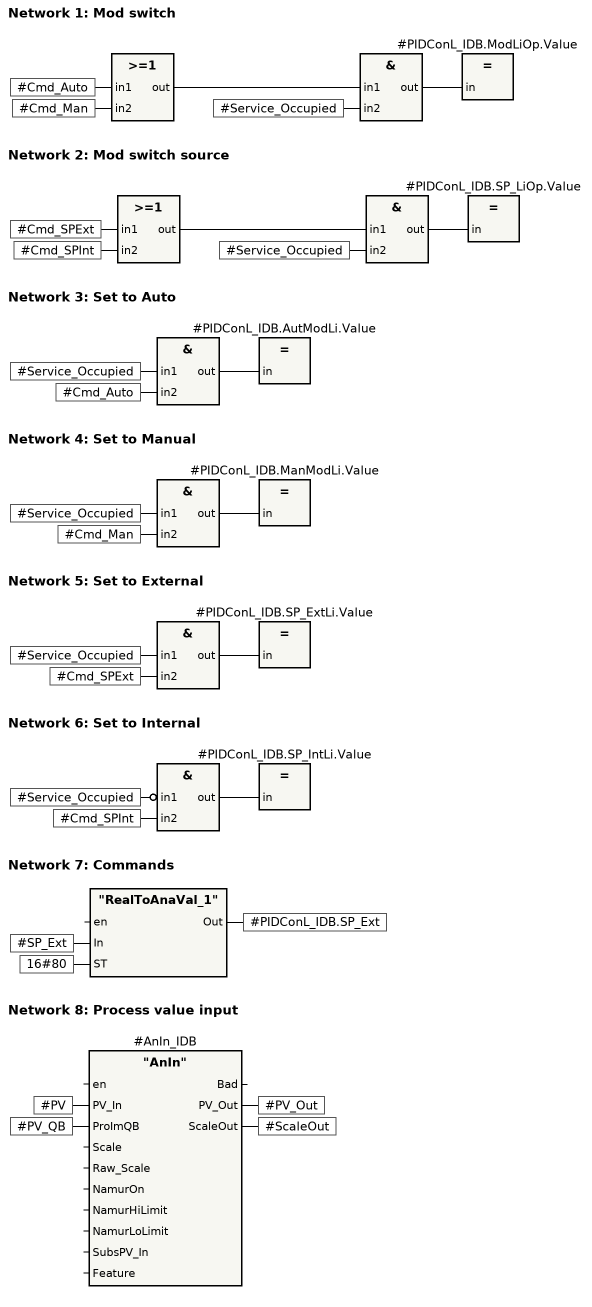
   #PIDConL_IDB.ModLiOp.Value := (#Cmd_Auto OR #Cmd_Man) AND #Service_Occupied;
END_REGION

REGION Network 2: Mod switch source
   #PIDConL_IDB.SP_LiOp.Value := (#Cmd_SPExt OR #Cmd_SPInt) AND #Service_Occupied;
END_REGION

REGION Network 3: Set to Auto
   #PIDConL_IDB.AutModLi.Value := #Service_Occupied AND #Cmd_Auto;
END_REGION

REGION Network 4: Set to Manual
   #PIDConL_IDB.ManModLi.Value := #Service_Occupied AND #Cmd_Man;
END_REGION

REGION Network 5: Set to External
   #PIDConL_IDB.SP_ExtLi.Value := #Service_Occupied AND #Cmd_SPExt;
END_REGION

REGION Network 6: Set to Internal
   #PIDConL_IDB.SP_IntLi.Value := NOT #Service_Occupied AND #Cmd_SPInt;
END_REGION

REGION Network 7: Commands
   "RealToAnaVal_1"(In := #SP_Ext, ST := 16#80, Out => #PIDConL_IDB.SP_Ext);
END_REGION

REGION Network 8: Process value input
   #AnIn_IDB(PV_In := #PV, ProImQB := #PV_QB, PV_Out => #PV_Out, ScaleOut => #ScaleOut);   // "AnIn"
END_REGION

REGION Network 9: CSF
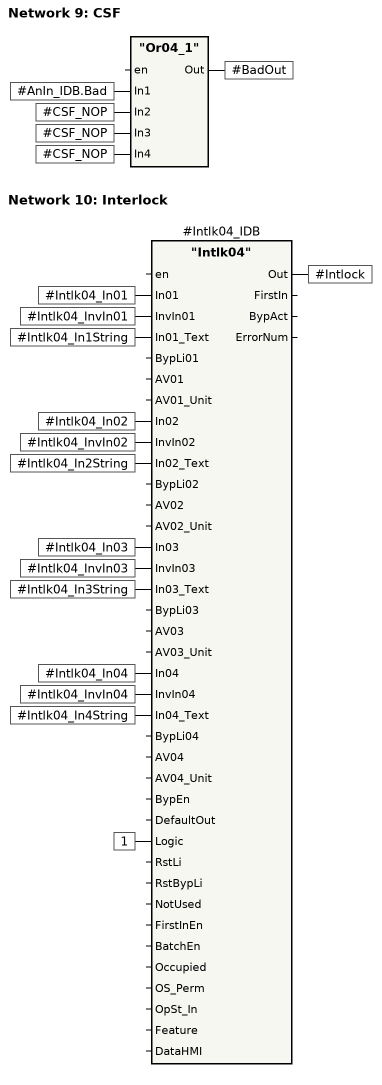
   "Or04_1"(In1 := #AnIn_IDB.Bad, In2 := #CSF_NOP, In3 := #CSF_NOP, In4 := #CSF_NOP, Out => #BadOut);
END_REGION

REGION Network 10: Interlock
   #Intlk04_IDB(In01 := #Intlk04_In01,   // "Intlk04"
                InvIn01 := #Intlk04_InvIn01,
                In01_Text := #Intlk04_In1String,
                In02 := #Intlk04_In02,
                InvIn02 := #Intlk04_InvIn02,
                In02_Text := #Intlk04_In2String,
                In03 := #Intlk04_In03,
                InvIn03 := #Intlk04_InvIn03,
                In03_Text := #Intlk04_In3String,
                In04 := #Intlk04_In04,
                InvIn04 := #Intlk04_InvIn04,
                In04_Text := #Intlk04_In4String,
                Logic := 1,
                Out => #Intlock);
END_REGION

REGION Network 11: PIDCtrL / PIDConL
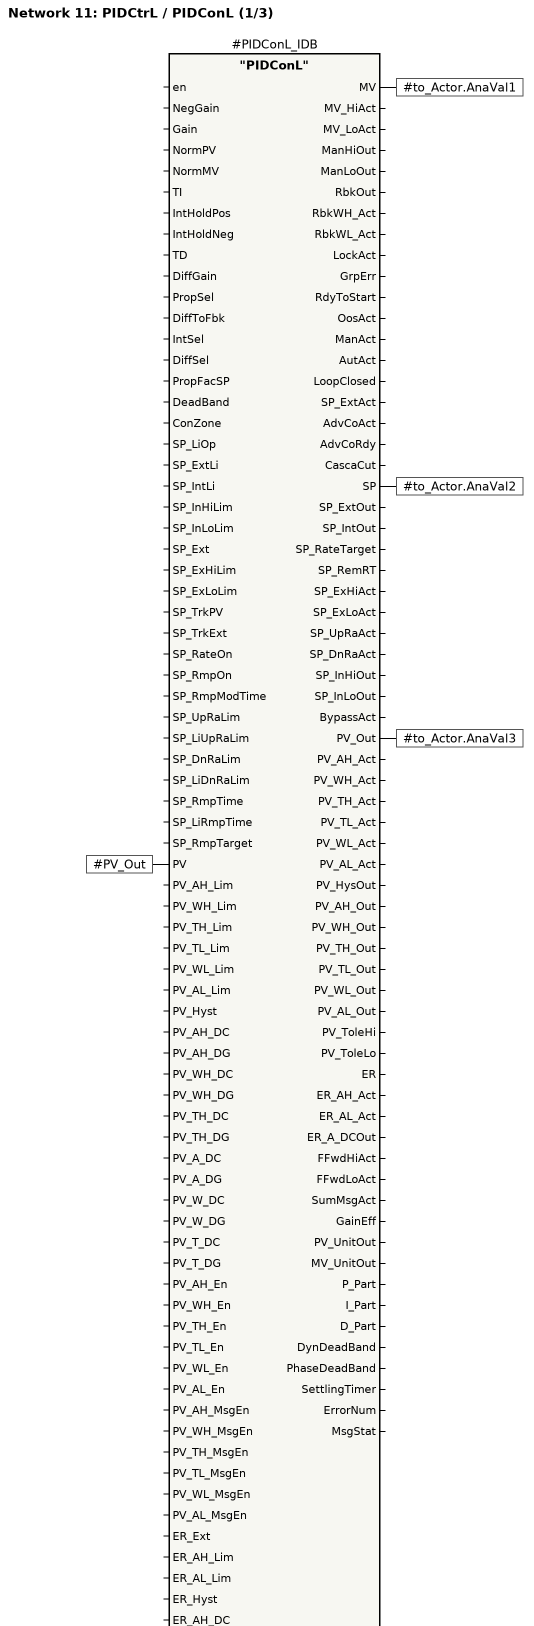
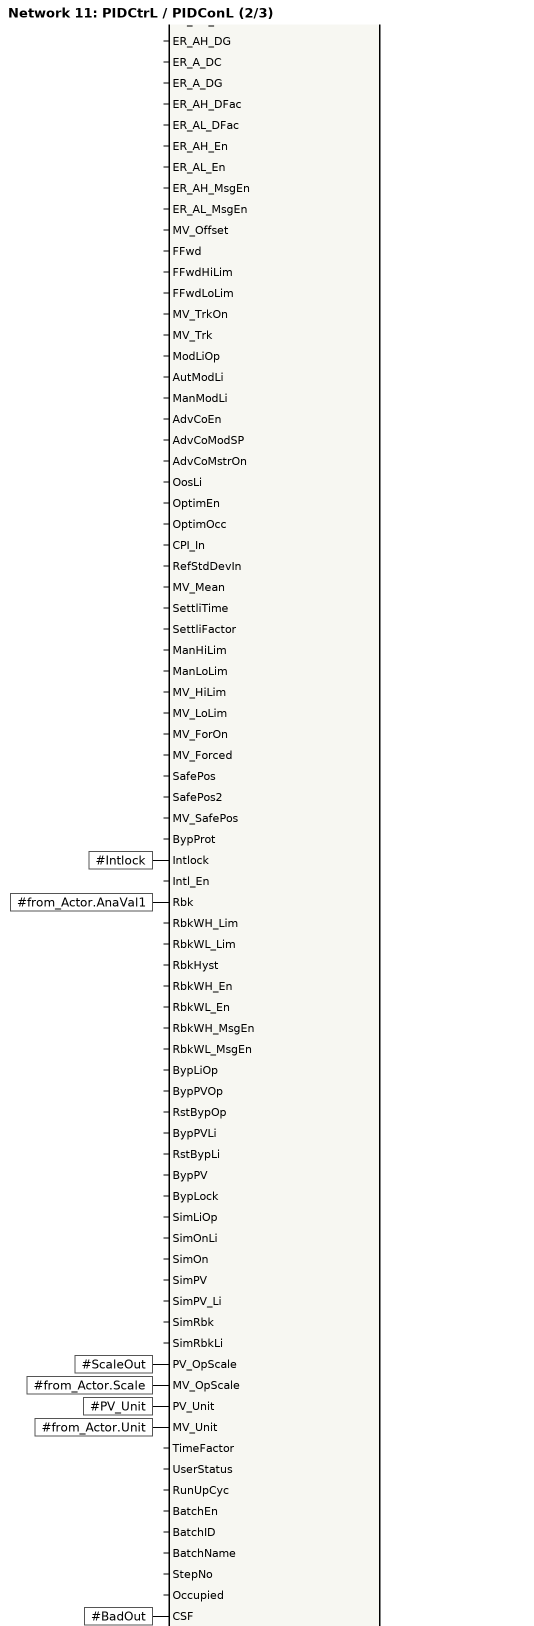
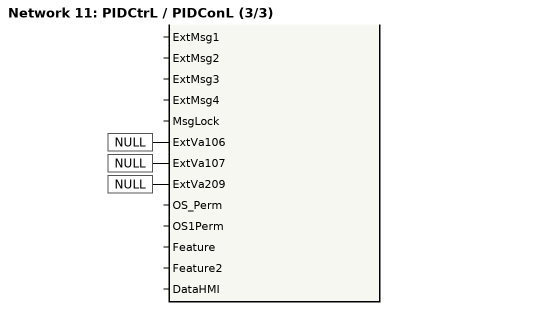
   #PIDConL_IDB(PV := #PV_Out,   // "PIDConL"
                Intlock := #Intlock,
                Rbk := #from_Actor.AnaVal1,
                PV_OpScale := #ScaleOut,
                MV_OpScale := #from_Actor.Scale,
                PV_Unit := #PV_Unit,
                MV_Unit := #from_Actor.Unit,
                CSF := #BadOut,
                ExtVa106 := NULL,
                ExtVa107 := NULL,
                ExtVa209 := NULL,
                MV => #to_Actor.AnaVal1,
                SP => #to_Actor.AnaVal2,
                PV_Out => #to_Actor.AnaVal3);
END_REGION

REGION Network 12: MTPPIDCtrl
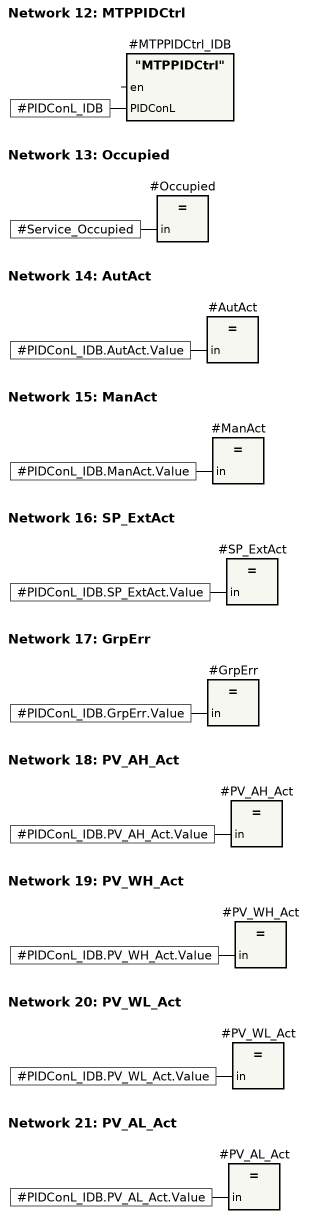
   #MTPPIDCtrl_IDB(PIDConL := #PIDConL_IDB);   // "MTPPIDCtrl"
END_REGION

REGION Network 13: Occupied
   #Occupied := #Service_Occupied;
END_REGION

REGION Network 14: AutAct
   #AutAct := #PIDConL_IDB.AutAct.Value;
END_REGION

REGION Network 15: ManAct
   #ManAct := #PIDConL_IDB.ManAct.Value;
END_REGION

REGION Network 16: SP_ExtAct
   #SP_ExtAct := #PIDConL_IDB.SP_ExtAct.Value;
END_REGION

REGION Network 17: GrpErr
   #GrpErr := #PIDConL_IDB.GrpErr.Value;
END_REGION

REGION Network 18: PV_AH_Act
   #PV_AH_Act := #PIDConL_IDB.PV_AH_Act.Value;
END_REGION

REGION Network 19: PV_WH_Act
   #PV_WH_Act := #PIDConL_IDB.PV_WH_Act.Value;
END_REGION

REGION Network 20: PV_WL_Act
   #PV_WL_Act := #PIDConL_IDB.PV_WL_Act.Value;
END_REGION

REGION Network 21: PV_AL_Act
   #PV_AL_Act := #PIDConL_IDB.PV_AL_Act.Value;
END_REGION
END_FUNCTION_BLOCK

FUNCTION "RealToAnaVal_1" : Void   // FC16, SCL
{ S7_Optimized_Access := 'TRUE' }
// stored: SetENOAutomatically false
   VAR_INPUT
      In : Real;
      ST : Byte;
   END_VAR
   VAR_OUTPUT
      Out : "AnaVal";
   END_VAR
BEGIN
   #Out.ST := #ST;
   #Out.Value := #In;
END_FUNCTION

FUNCTION "FIT100" : Void   // FC4, FBD
{ S7_Optimized_Access := 'TRUE' }
// stored: SetENOAutomatically false
   VAR_TEMP
      Temp : "DigVal";
      Temp_1 : "DigVal";
   END_VAR
BEGIN

REGION Network 1: MonAnL
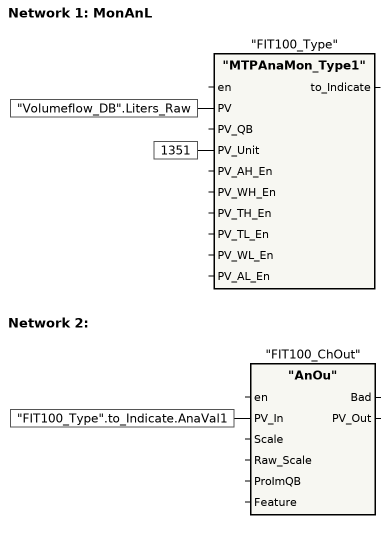
   "FIT100_Type"(PV := "Volumeflow_DB".Liters_Raw, PV_Unit := 1351);   // "MTPAnaMon_Type1"
END_REGION

REGION Network 2
   "FIT100_ChOut"(PV_In := "FIT100_Type".to_Indicate.AnaVal1);   // "AnOu"
END_REGION
END_FUNCTION

FUNCTION_BLOCK "MTPAnaMon_Type1"   // FB15, FBD
{ S7_Optimized_Access := 'TRUE' }
// stored: MemoryReserve 100, SetENOAutomatically false
   VAR_INPUT
      PV { ExternalAccessible := 'False'; ExternalVisible := 'False'; ExternalWritable := 'False'} : Word;
      PV_QB { ExternalAccessible := 'False'; ExternalVisible := 'False'; ExternalWritable := 'False'} : Bool := true;
      PV_Unit { ExternalAccessible := 'False'; ExternalVisible := 'False'; ExternalWritable := 'False'} : Int := 1001;
      PV_AH_En { ExternalAccessible := 'False'; ExternalVisible := 'False'; ExternalWritable := 'False'} : Bool := true;
      PV_WH_En { ExternalAccessible := 'False'; ExternalVisible := 'False'; ExternalWritable := 'False'} : Bool := true;
      PV_TH_En { ExternalAccessible := 'False'; ExternalVisible := 'False'; ExternalWritable := 'False'} : Bool;
      PV_TL_En { ExternalAccessible := 'False'; ExternalVisible := 'False'; ExternalWritable := 'False'} : Bool;
      PV_WL_En { ExternalAccessible := 'False'; ExternalVisible := 'False'; ExternalWritable := 'False'} : Bool := true;
      PV_AL_En { ExternalAccessible := 'False'; ExternalVisible := 'False'; ExternalWritable := 'False'} : Bool := true;
   END_VAR
   VAR_OUTPUT
      to_Indicate { ExternalAccessible := 'False'; ExternalVisible := 'False'; ExternalWritable := 'False'} : "StruCm";
   END_VAR
   VAR
      AnIn_IDB { ExternalAccessible := 'False'; ExternalVisible := 'False'; ExternalWritable := 'False'} : "AnIn";
      MonAnL_IDB : "MonAnL";
      MTPAnaMon_IDB { ExternalVisible := 'False'; S7_SetPoint := 'True'} : "MTPAnaMon";
   END_VAR
   VAR_TEMP
      PV_Out : "AnaVal";
      CSF_NOP : "DigVal";
      BadAnIn : "DigVal";
      BadOut : "DigVal";
      ScaleOut : "ScaVal";
   END_VAR
   VAR_TEMP   // added for the SCL form of the ladder/FBD networks
      _w1 : Bool;
   END_VAR
BEGIN

REGION Network 1: Convert / Init
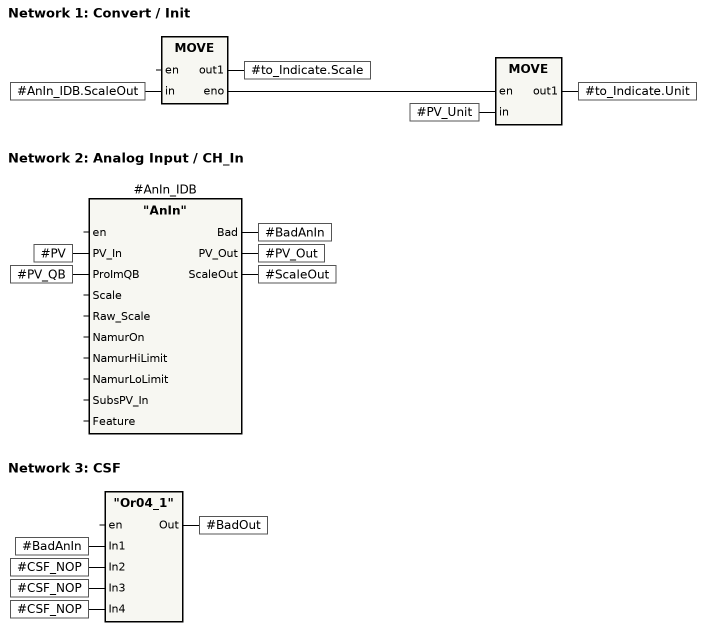
   #to_Indicate.Scale := #AnIn_IDB.ScaleOut;
   #to_Indicate.Unit := #PV_Unit;
END_REGION

REGION Network 2: Analog Input / CH_In
   #AnIn_IDB(PV_In := #PV, ProImQB := #PV_QB, Bad => #BadAnIn, PV_Out => #PV_Out, ScaleOut => #ScaleOut);   // "AnIn"
END_REGION

REGION Network 3: CSF
   "Or04_1"(In1 := #BadAnIn, In2 := #CSF_NOP, In3 := #CSF_NOP, In4 := #CSF_NOP, Out => #BadOut);
END_REGION

REGION Network 4: MonAnL
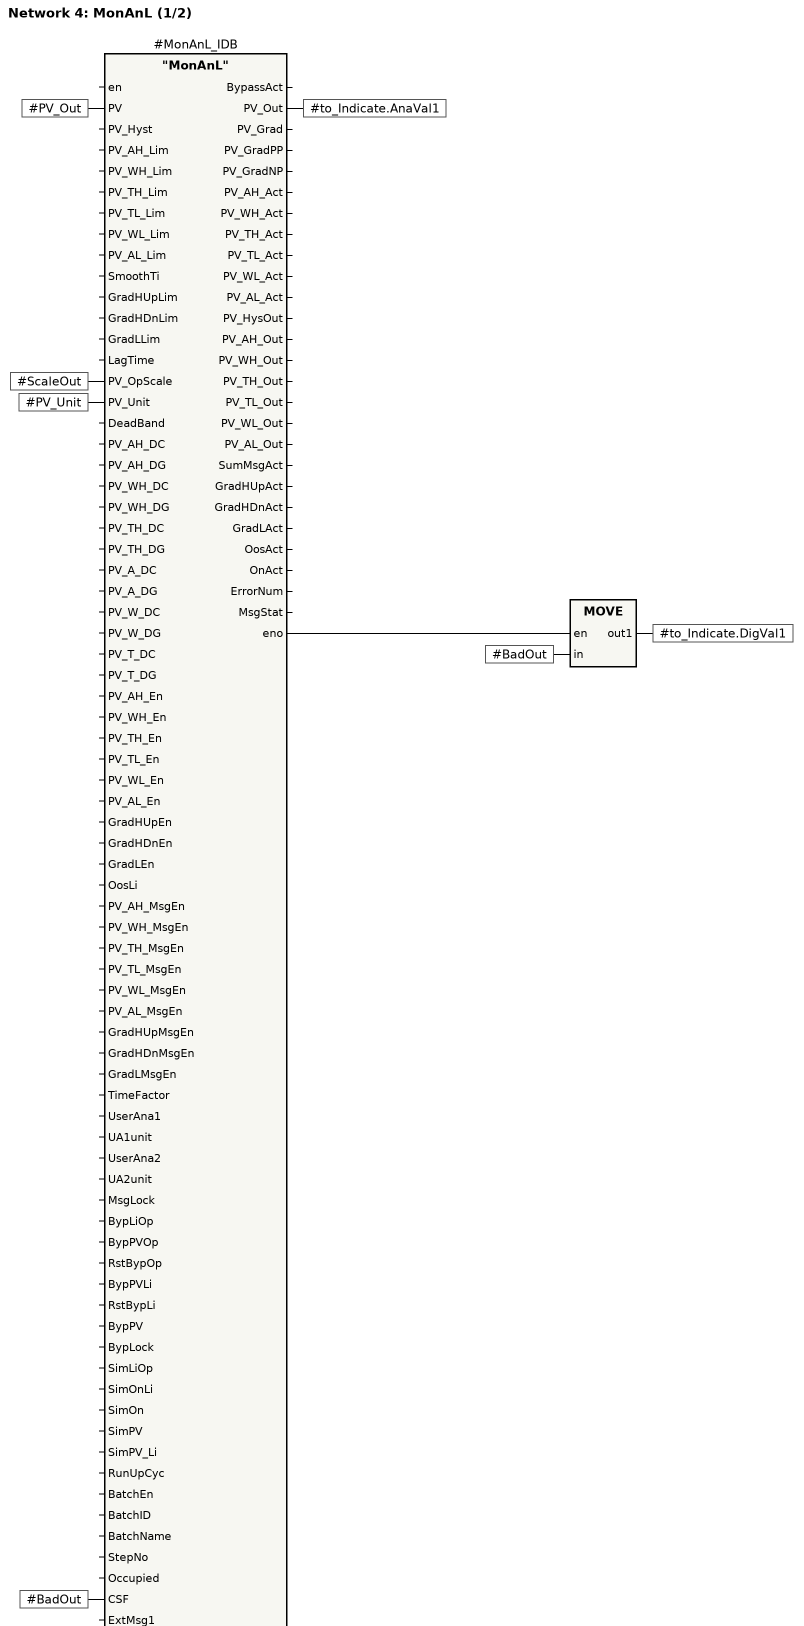
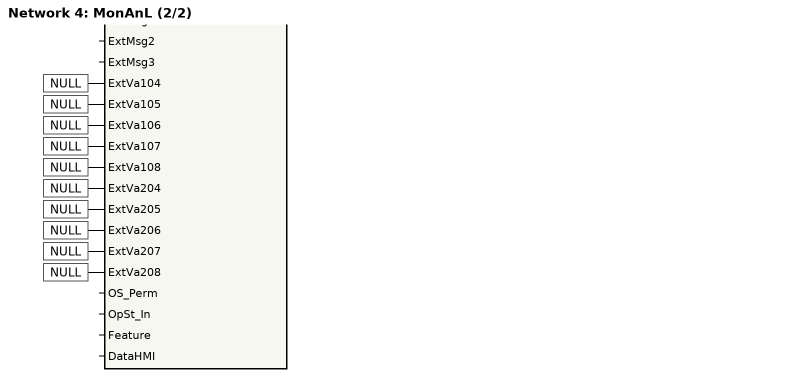
   #MonAnL_IDB(PV := #PV_Out,   // "MonAnL"
               PV_OpScale := #ScaleOut,
               PV_Unit := #PV_Unit,
               CSF := #BadOut,
               ExtVa104 := NULL,
               ExtVa105 := NULL,
               ExtVa106 := NULL,
               ExtVa107 := NULL,
               ExtVa108 := NULL,
               ExtVa204 := NULL,
               ExtVa205 := NULL,
               ExtVa206 := NULL,
               ExtVa207 := NULL,
               ExtVa208 := NULL,
               PV_Out => #to_Indicate.AnaVal1,
               ENO => #_w1);
   IF #_w1 THEN #to_Indicate.DigVal1 := #BadOut; END_IF;
END_REGION

REGION Network 5: MTP / MTP Connector block
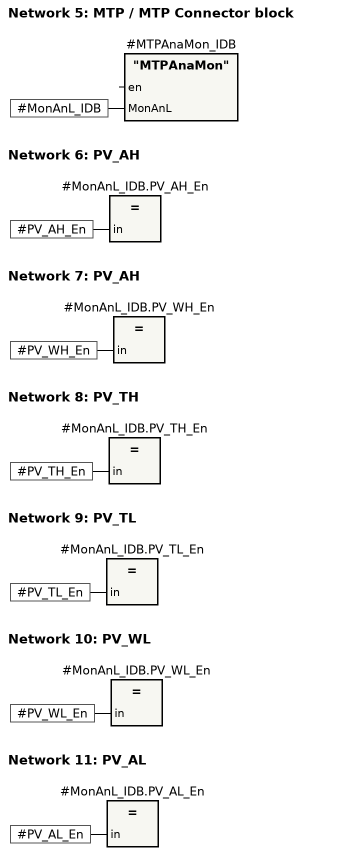
   #MTPAnaMon_IDB(MonAnL := #MonAnL_IDB);   // "MTPAnaMon"
END_REGION

REGION Network 6: PV_AH
   #MonAnL_IDB.PV_AH_En := #PV_AH_En;
END_REGION

REGION Network 7: PV_AH
   #MonAnL_IDB.PV_WH_En := #PV_WH_En;
END_REGION

REGION Network 8: PV_TH
   #MonAnL_IDB.PV_TH_En := #PV_TH_En;
END_REGION

REGION Network 9: PV_TL
   #MonAnL_IDB.PV_TL_En := #PV_TL_En;
END_REGION

REGION Network 10: PV_WL
   #MonAnL_IDB.PV_WL_En := #PV_WL_En;
END_REGION

REGION Network 11: PV_AL
   #MonAnL_IDB.PV_AL_En := #PV_AL_En;
END_REGION
END_FUNCTION_BLOCK

FUNCTION "FIT100_Liter" : Void   // FC15, FBD
{ S7_Optimized_Access := 'TRUE' }
// stored: SetENOAutomatically false
BEGIN

REGION Network 1: MonAnL
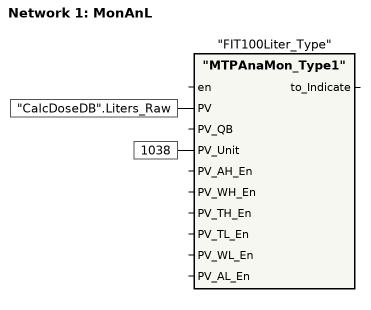
   "FIT100Liter_Type"(PV := "CalcDoseDB".Liters_Raw, PV_Unit := 1038);   // "MTPAnaMon_Type1"
END_REGION
END_FUNCTION

FUNCTION "LAH100" : Void   // FC8, FBD
{ S7_Optimized_Access := 'TRUE' }
// stored: SetENOAutomatically false
BEGIN

REGION Network 1: MonDiL
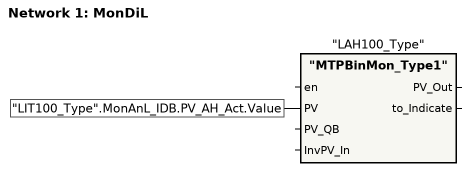
   "LAH100_Type"(PV := "LIT100_Type".MonAnL_IDB.PV_AH_Act.Value);   // "MTPBinMon_Type1"
END_REGION
END_FUNCTION

FUNCTION_BLOCK "MTPBinMon_Type1"   // FB16, FBD
{ S7_Optimized_Access := 'TRUE' }
// stored: MemoryReserve 100, SetENOAutomatically false
   VAR_INPUT
      PV { ExternalAccessible := 'False'; ExternalVisible := 'False'; ExternalWritable := 'False'} : Bool;
      PV_QB { ExternalAccessible := 'False'; ExternalVisible := 'False'; ExternalWritable := 'False'} : Bool := true;
      InvPV_In { ExternalAccessible := 'False'; ExternalVisible := 'False'; ExternalWritable := 'False'} : Bool;
   END_VAR
   VAR_OUTPUT
      PV_Out { ExternalAccessible := 'False'; ExternalVisible := 'False'; ExternalWritable := 'False'} : Bool;
      to_Indicate { ExternalAccessible := 'False'; ExternalVisible := 'False'; ExternalWritable := 'False'} : "StruCm";
   END_VAR
   VAR
      DiIn_IDB { ExternalAccessible := 'False'; ExternalVisible := 'False'; ExternalWritable := 'False'} : "DiIn";
      MonDiL_IDB { S7_SetPoint := 'True'} : "MonDiL";
      MTPBinMon_IDB { ExternalVisible := 'False'; S7_SetPoint := 'True'} : "MTPBinMon";
   END_VAR
   VAR_TEMP
      PV_Out_Temp : "DigVal";
      CSF_NOP : "DigVal";
      BadDiIn : "DigVal";
      BadOut : "DigVal";
   END_VAR
   VAR_TEMP   // added for the SCL form of the ladder/FBD networks
      _w1 : Bool;
   END_VAR
BEGIN

REGION Network 1: Analog Input
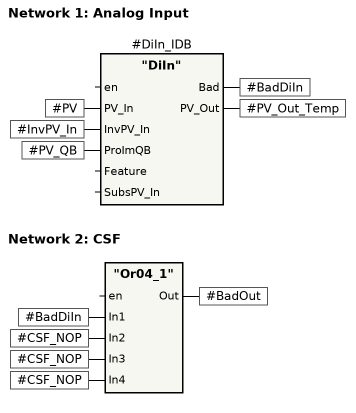
   #DiIn_IDB(PV_In := #PV, InvPV_In := #InvPV_In, ProImQB := #PV_QB, Bad => #BadDiIn, PV_Out => #PV_Out_Temp);   // "DiIn"
END_REGION

REGION Network 2: CSF
   "Or04_1"(In1 := #BadDiIn, In2 := #CSF_NOP, In3 := #CSF_NOP, In4 := #CSF_NOP, Out => #BadOut);
END_REGION

REGION Network 3: MonAnL
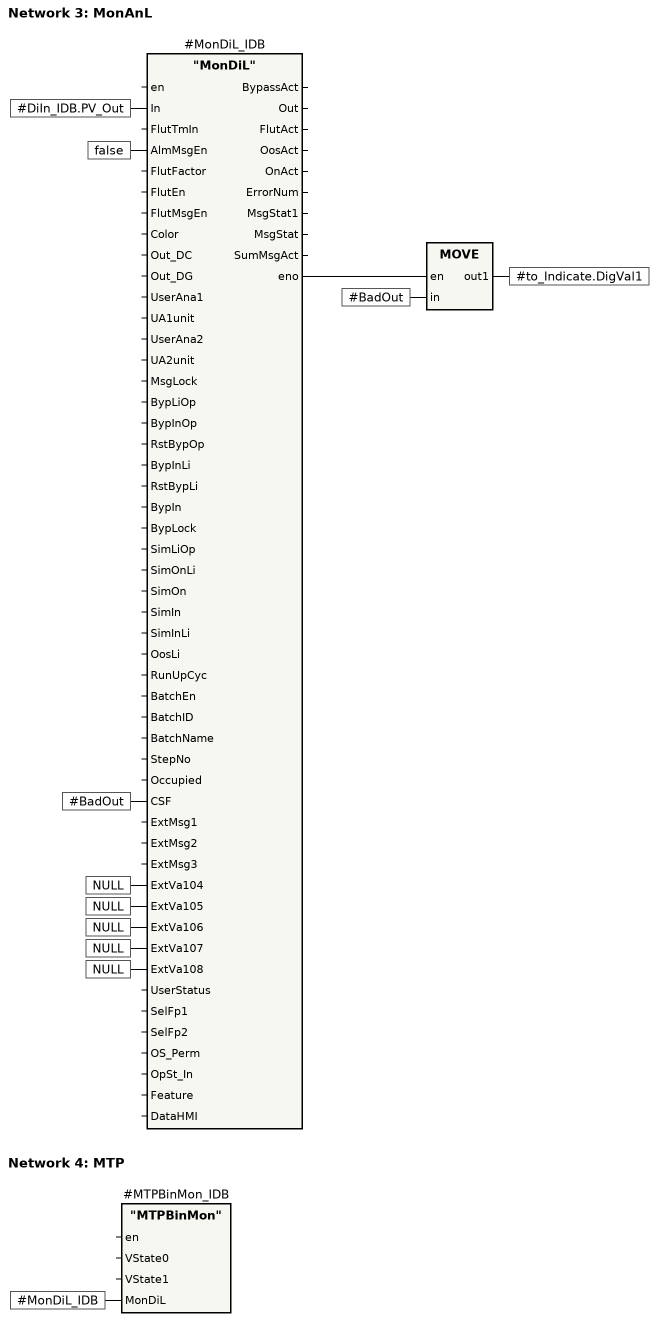
   #MonDiL_IDB(In := #DiIn_IDB.PV_Out,   // "MonDiL"
               AlmMsgEn := false,
               CSF := #BadOut,
               ExtVa104 := NULL,
               ExtVa105 := NULL,
               ExtVa106 := NULL,
               ExtVa107 := NULL,
               ExtVa108 := NULL,
               ENO => #_w1);
   IF #_w1 THEN #to_Indicate.DigVal1 := #BadOut; END_IF;
END_REGION

REGION Network 4: MTP
   #MTPBinMon_IDB(MonDiL := #MonDiL_IDB);   // "MTPBinMon"
END_REGION

REGION Network 5
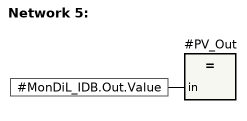
   #PV_Out := #MonDiL_IDB.Out.Value;
END_REGION
END_FUNCTION_BLOCK

FUNCTION "LAL100" : Void   // FC7, FBD
{ S7_Optimized_Access := 'TRUE' }
// stored: SetENOAutomatically false
BEGIN

REGION Network 1: MonDiL
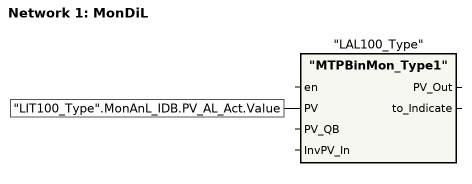
   "LAL100_Type"(PV := "LIT100_Type".MonAnL_IDB.PV_AL_Act.Value);   // "MTPBinMon_Type1"
END_REGION
END_FUNCTION

FUNCTION "LIT100" : Void   // FC6, FBD
{ S7_Optimized_Access := 'TRUE' }
// stored: SetENOAutomatically false
BEGIN

REGION Network 1: Tank level
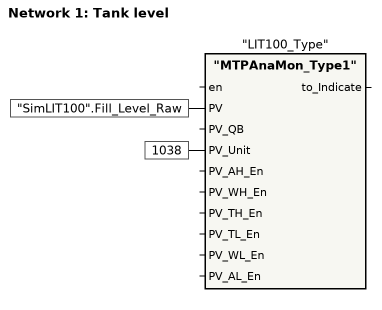
   "LIT100_Type"(PV := "SimLIT100".Fill_Level_Raw, PV_Unit := 1038);   // "MTPAnaMon_Type1"
END_REGION
END_FUNCTION

FUNCTION "P100" : Void   // FC2, FBD
{ S7_Optimized_Access := 'TRUE' }
// stored: SetENOAutomatically false
   VAR_TEMP
      Temp : "DigVal";
      Temp_1 : "DigVal";
      Temp_3 : "DigVal";
      Temp_2 : "DigVal";
      Temp_Error : "DigVal";
      In03 : "DigVal";
      State : "Service_States";
      FbkRun : "DigVal";
      StopAut : Bool;
   END_VAR
   VAR_TEMP   // added for the SCL form of the ladder/FBD networks
      _w1 : Bool;
   END_VAR
BEGIN

REGION Network 1: simulate Fbk Error
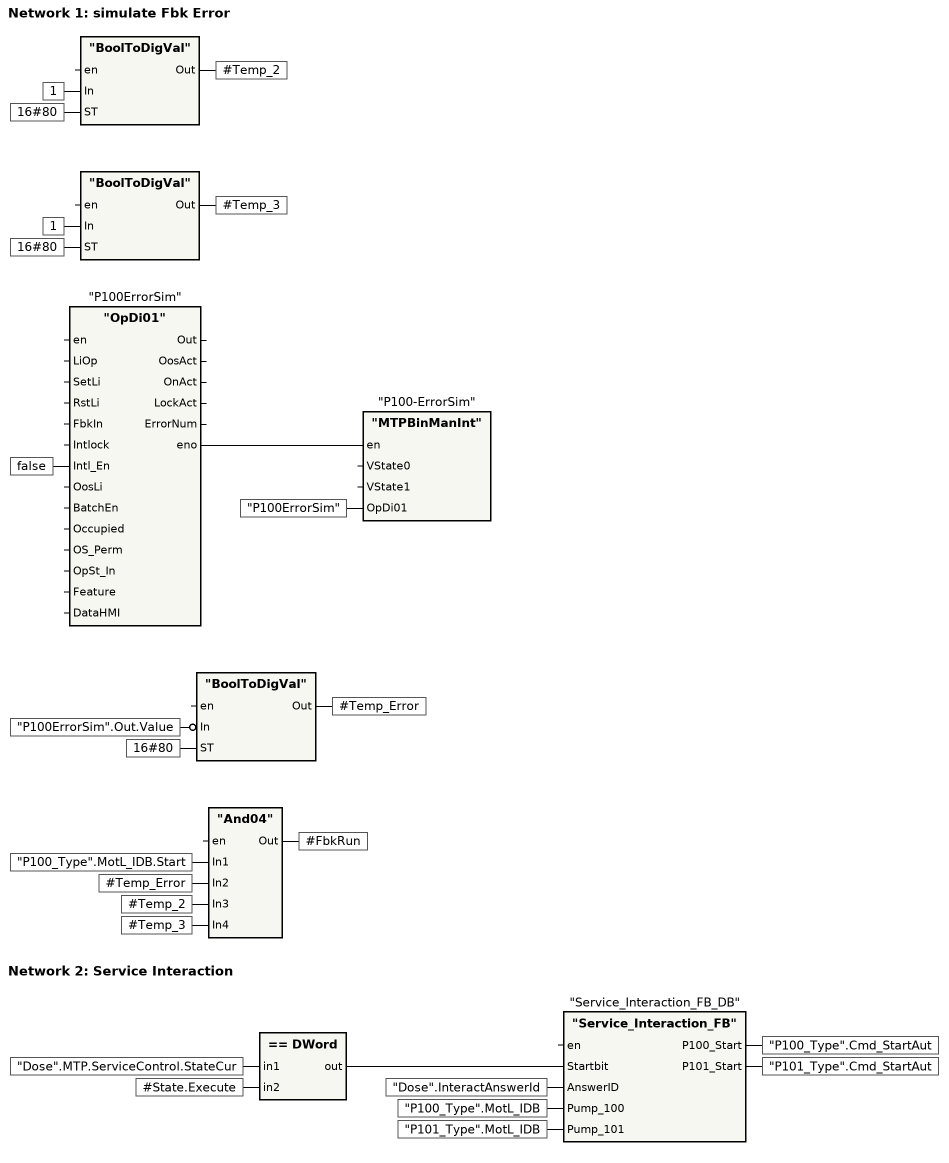
   "BoolToDigVal"(In := 1, ST := 16#80, Out => #Temp_2);
   "BoolToDigVal"(In := 1, ST := 16#80, Out => #Temp_3);
   "P100ErrorSim"(Intl_En := false, ENO => #_w1);   // "OpDi01"
   IF #_w1 THEN
       "P100-ErrorSim"(OpDi01 := "P100ErrorSim");   // "MTPBinManInt"
   END_IF;
   "BoolToDigVal"(In := NOT "P100ErrorSim".Out.Value, ST := 16#80, Out => #Temp_Error);
   "And04"(In1 := "P100_Type".MotL_IDB.Start,
           In2 := #Temp_Error,
           In3 := #Temp_2,
           In4 := #Temp_3,
           Out => #FbkRun);
END_REGION

REGION Network 2: Service Interaction
   "Service_Interaction_FB_DB"(Startbit := "Dose".MTP.ServiceControl.StateCur = #State.Execute,   // "Service_Interaction_FB"
                           AnswerID := "Dose".InteractAnswerId,
                           Pump_100 := "P100_Type".MotL_IDB,
                           Pump_101 := "P101_Type".MotL_IDB,
                           P100_Start => "P100_Type".Cmd_StartAut,
                           P101_Start => "P101_Type".Cmd_StartAut);
END_REGION

REGION Network 3: Pump interconnections
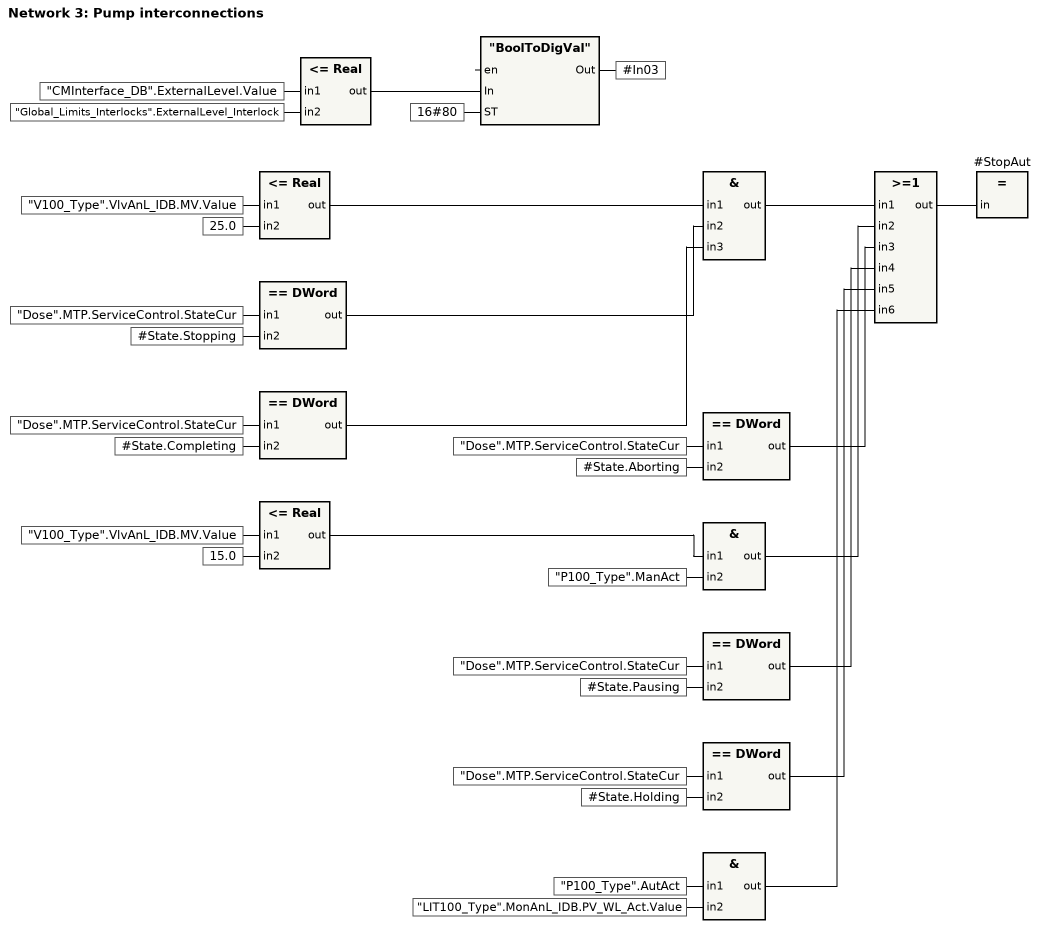
   "BoolToDigVal"(In := "CMInterface_DB".ExternalLevel.Value <= "Global_Limits_Interlocks".ExternalLevel_Interlock,
                  ST := 16#80,
                  Out => #In03);
   #StopAut := (("V100_Type".VlvAnL_IDB.MV.Value <= 25.0) AND ("Dose".MTP.ServiceControl.StateCur = #State.Stopping) AND ("Dose".MTP.ServiceControl.StateCur = #State.Completing)) OR (("V100_Type".VlvAnL_IDB.MV.Value <= 15.0) AND "P100_Type".ManAct) OR ("Dose".MTP.ServiceControl.StateCur = #State.Aborting) OR ("Dose".MTP.ServiceControl.StateCur = #State.Pausing) OR ("Dose".MTP.ServiceControl.StateCur = #State.Holding) OR ("P100_Type".AutAct AND "LIT100_Type".MonAnL_IDB.PV_WL_Act.Value);
END_REGION

REGION Network 4: MotL
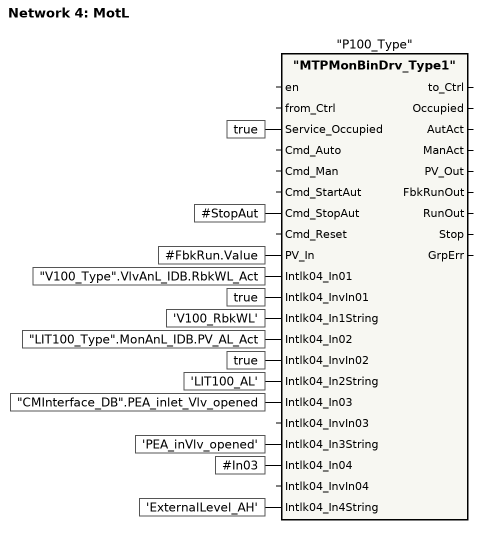
   "P100_Type"(Service_Occupied := true,   // "MTPMonBinDrv_Type1"
               Cmd_StopAut := #StopAut,
               PV_In := #FbkRun.Value,
               Intlk04_In01 := "V100_Type".VlvAnL_IDB.RbkWL_Act,
               Intlk04_InvIn01 := true,
               Intlk04_In1String := 'V100_RbkWL',
               Intlk04_In02 := "LIT100_Type".MonAnL_IDB.PV_AL_Act,
               Intlk04_InvIn02 := true,
               Intlk04_In2String := 'LIT100_AL',
               Intlk04_In03 := "CMInterface_DB".PEA_inlet_Vlv_opened,
               Intlk04_In3String := 'PEA_inVlv_opened',
               Intlk04_In04 := #In03,
               Intlk04_In4String := 'ExternalLevel_AH');
END_REGION
END_FUNCTION

FUNCTION_BLOCK "Service_Interaction_FB"   // FB6, SCL
{ S7_Optimized_Access := 'TRUE' }
// stored: MemoryReserve 100, SetENOAutomatically false
   VAR_INPUT
      Startbit { ExternalAccessible := 'False'; ExternalVisible := 'False'; ExternalWritable := 'False'} : Bool;
      AnswerID { ExternalAccessible := 'False'; ExternalVisible := 'False'; ExternalWritable := 'False'} : DWord;
   END_VAR
   VAR_OUTPUT
      P100_Start : Bool;
      P101_Start : Bool;
   END_VAR
   VAR_IN_OUT
      Pump_100 : "MotL";
      Pump_101 : "MotL";
   END_VAR
   VAR_TEMP
      State : "Service_States";
   END_VAR
BEGIN
   //if positive edge, then trigger service interaction (set Question and info text)
   IF #Startbit AND NOT #Pump_100.Run.Value AND NOT #Pump_101.Run.Value THEN
       "Dose".InteractAddInfoLi := 'Select the available Pump for the operation';
       "Dose".InteractQuestionIdLi := 1;
   END_IF;

   //if answer ID 1 or 3 is selected, start pump_100
   IF ((#AnswerID = 1 OR #AnswerID = 3) AND #Startbit) THEN
       #P100_Start := True;
   END_IF;
   //if answer ID 2 or 3 is selected, start pump_101
   IF ((#AnswerID = 2 OR #AnswerID = 3) AND #Startbit) THEN
       #P101_Start := True;
   END_IF;

   //if answer ID 0 or service in state stopping/resetting/aborting/completing then reset question ID and info
   IF (#AnswerID <> 0 AND #Startbit) OR "Dose".MTP.ServiceControl.StateCur <> #State.Execute THEN
       "Dose".InteractQuestionIdLi := 0;
       "Dose".InteractAddInfoLi := '';
   END_IF;

   //reset start aut of pumps, if no positive edge
   IF NOT #Startbit AND (#Pump_100.Run.Value = True OR #Pump_101.Run.Value = True) THEN
       #P100_Start := false;
       #P101_Start := false;
   END_IF;
END_FUNCTION_BLOCK

FUNCTION_BLOCK "MTPMonBinDrv_Type1"   // FB13, FBD
{ S7_Optimized_Access := 'TRUE' }
// stored: MemoryReserve 100, SetENOAutomatically false
   VAR_INPUT
      from_Ctrl { ExternalAccessible := 'False'; ExternalVisible := 'False'; ExternalWritable := 'False'} : "StruCm";
      Service_Occupied { ExternalAccessible := 'False'; ExternalVisible := 'False'; ExternalWritable := 'False'} : Bool;
      Cmd_Auto { ExternalAccessible := 'False'; ExternalVisible := 'False'; ExternalWritable := 'False'} : Bool;
      Cmd_Man { ExternalAccessible := 'False'; ExternalVisible := 'False'; ExternalWritable := 'False'} : Bool;
      Cmd_StartAut { ExternalAccessible := 'False'; ExternalVisible := 'False'; ExternalWritable := 'False'} : Bool;
      Cmd_StopAut { ExternalAccessible := 'False'; ExternalVisible := 'False'; ExternalWritable := 'False'} : Bool;
      Cmd_Reset { ExternalAccessible := 'False'; ExternalVisible := 'False'; ExternalWritable := 'False'} : Bool;
      PV_In : Bool;
      Intlk04_In01 { ExternalAccessible := 'False'; ExternalVisible := 'False'; ExternalWritable := 'False'} : "DigVal";
      Intlk04_InvIn01 : Bool;
      Intlk04_In1String : String;
      Intlk04_In02 { ExternalAccessible := 'False'; ExternalVisible := 'False'; ExternalWritable := 'False'} : "DigVal";
      Intlk04_InvIn02 : Bool;
      Intlk04_In2String { ExternalAccessible := 'False'; ExternalVisible := 'False'; ExternalWritable := 'False'} : String;
      Intlk04_In03 { ExternalAccessible := 'False'; ExternalVisible := 'False'; ExternalWritable := 'False'} : "DigVal";
      Intlk04_InvIn03 : Bool;
      Intlk04_In3String { ExternalAccessible := 'False'; ExternalVisible := 'False'; ExternalWritable := 'False'} : String;
      Intlk04_In04 { ExternalAccessible := 'False'; ExternalVisible := 'False'; ExternalWritable := 'False'} : "DigVal";
      Intlk04_InvIn04 : Bool;
      Intlk04_In4String { ExternalAccessible := 'False'; ExternalVisible := 'False'; ExternalWritable := 'False'} : String;
   END_VAR
   VAR_OUTPUT
      to_Ctrl { ExternalAccessible := 'False'; ExternalVisible := 'False'; ExternalWritable := 'False'} : "StruCm";
      Occupied { ExternalAccessible := 'False'; ExternalVisible := 'False'; ExternalWritable := 'False'} : Bool;   // Occupied by a Service procedure
      AutAct { ExternalAccessible := 'False'; ExternalVisible := 'False'; ExternalWritable := 'False'} : Bool;
      ManAct { ExternalAccessible := 'False'; ExternalVisible := 'False'; ExternalWritable := 'False'} : Bool;
      PV_Out { ExternalAccessible := 'False'; ExternalVisible := 'False'; ExternalWritable := 'False'} : Bool;
      FbkRunOut : Bool;
      RunOut : Bool;
      Stop { ExternalAccessible := 'False'; ExternalVisible := 'False'; ExternalWritable := 'False'} : Bool;
      GrpErr { ExternalAccessible := 'False'; ExternalVisible := 'False'; ExternalWritable := 'False'} : Bool;
   END_VAR
   VAR
      ChOut { S7_SetPoint := 'True'} : "DiOu";
      DiChIn { S7_SetPoint := 'True'} : "DiIn";
      Intlk04_IDB : "Intlk04";
      MotL_IDB { S7_SetPoint := 'True'} : "MotL";
      MTPMonBinDrv_IDB { ExternalVisible := 'False'; S7_SetPoint := 'True'} : "MTPMonBinDrv";
   END_VAR
   VAR_TEMP
      Intlock : "DigVal";
      CSF_NOP : "DigVal";
      BadOut : "DigVal";
      InverterBad : "DigVal";
      FbkRun : "DigVal";
   END_VAR
   // Intlk04_In01.Value := true;
   // Intlk04_In02.Value := true;
   // Intlk04_In03.Value := true;
   // Intlk04_In04.Value := true;
BEGIN

REGION Network 1: Mod switch
